ABB RobotStudio station: Laboratorio1Ruiz.rspag

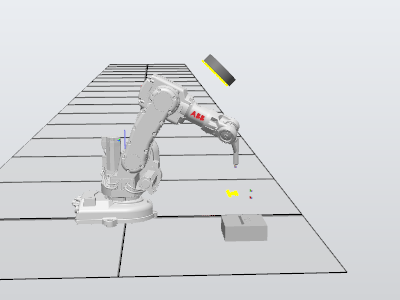
--- station ---
Station Laboratorio1 (saved by RobotStudio 25.5.11605.0)
Controller IRB140_6_81
  mechanical unit ROB_1: IRB140_6_81_C_03, 6 joints, base frame (0, 0, 0) mm
Layout (positions relative to the parent item):
  - IRB140_6_81_C_03 [mechanism, from %ABB.RobotStudio.Models.IRB140%\IRB140_6_81_C_G_03.rslib] at (0, 0, 0) mm; joint values [-0.1334, 0.4721, -0.017, 0.5827, 0.9537, -1.4192] (rad or m)
  - ToolLab1AlexaReyes [mechanism] at (588.01, -49.46, 449.3) mm, rotated rx 180 ry 30 rz -123.8 deg
      TCP ToolLab1AlexaReyes at (38.82, 1.24, 164.3) mm, rotated rx 0 ry 30 rz 0 deg
      links: Tool_3
  - Trayectorias2 [part] at (589.46, -613.7, 102.2) mm, rotated rx 0 ry 0 rz -90 deg, size 210 x 200 x 73 mm
  - Pieza_1 [part] at (-200, 0, 100) mm, rotated rx 0 ry 45 rz 0 deg, size 200 x 198.9 x 50 mm
  - SmartComponent_1 [smart component]
      signals: DI DI_04
      connections:
        LinearMover2.Executed -> LogicSRLatch.Reset
        LinearMover2.Executing -> LogicSRLatch.Set
        SmartComponent_1.DI_04 -> LinearMover2.Execute
    - LinearMover2 [smart component, from Components\LinearMover2.rslib]
        properties: Object=Trayectorias2; Direction=[0 0.001 0]; Distance=0.605; Duration=4.2; Reference=Global; ReferenceObject=(none)
  - SmartComponent_2 [smart component]
      signals: DI DI_05
      connections:
        SmartComponent_2.DI_05 -> LinearMover2_3.Execute
    - LinearMover2_3 [smart component, from Components\LinearMover2.rslib]
        properties: Object=Trayectorias2; Direction=[0 0.001 0]; Distance=0.605; Duration=4.2; Reference=Global; ReferenceObject=(none)
  - SmartComponent_3 [smart component]
      signals: DI DI_06
      connections:
        SmartComponent_3.DI_06 -> LinearMover2_5.Execute
    - LinearMover2_5 [smart component, from Components\LinearMover2.rslib]
        properties: Object=Trayectorias2; Direction=[0 -0.001 0]; Distance=1.21; Duration=8.4; Reference=Global; ReferenceObject=(none)
Attachment: ToolLab1AlexaReyes is attached to IRB140_6_81_C_03 / Link6
Station logic (signal -> signal, property => property):
  IRB140_6_81.DO_01 -> SmartComponent_1.DI_04
  IRB140_6_81.DO_02 -> SmartComponent_2.DI_05
  IRB140_6_81.DO_03 -> SmartComponent_3.DI_06

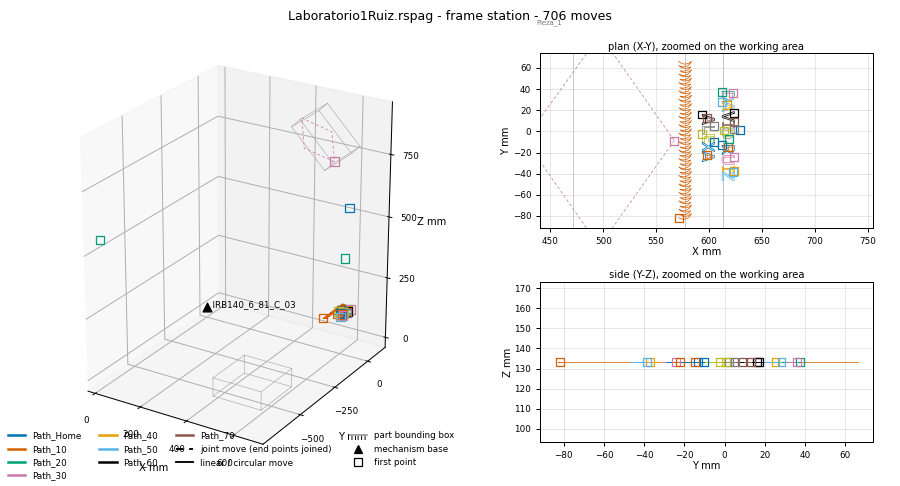
[picture p0: tool path of Laboratorio1Ruiz.rspag in frame station, 706 of 706 moves have a stored position in this frame; points joined in program order, loops and branches not executed]
--- Controller Data/IRB140_6_81/RAPID/TASK1/PROGMOD/Module1.mod ---
MODULE Module1
    PERS tooldata ToolLab1AlexaReyes:=[TRUE,[[38.819,1.24,164.297],[0.965925826,0,0.258819045,0]],[1,[0,0,1],[1,0,0,0],0,0,0]]; !CALIBRACIÓN VIRTUAL
    !PERS tooldata ToolLab1AlexaReyes:=[TRUE,[[37.2018,0.567088,156.366],[1,0,0,0]],[1,[0,0,0],[1,0,0,0],0,0,0]]; !CALIBRACIÓN FÍSICA
    CONST robtarget Target_Home:=[[629.167524851,1.24,563.73325724],[0.258819038,0,0.965925828,0],[0,-1,0,0],[9E+09,9E+09,9E+09,9E+09,9E+09,9E+09]];
    CONST robtarget Target_10:=[[118,32,0],[0.882142515,0,0,-0.470982573],[0,0,0,0],[9E+09,9E+09,9E+09,9E+09,9E+09,9E+09]];
    CONST robtarget Target_20:=[[115.336324555,30.849749419,0],[0.882142515,0,0,-0.470982573],[0,0,0,0],[9E+09,9E+09,9E+09,9E+09,9E+09,9E+09]];
    CONST robtarget Target_30:=[[112.437578714,30.725186884,0],[0.882142515,0,0,-0.470982573],[0,0,0,0],[9E+09,9E+09,9E+09,9E+09,9E+09,9E+09]];
    CONST robtarget Target_40:=[[109.685049159,31.642696736,0],[0.882142515,0,0,-0.470982573],[0,0,0,0],[9E+09,9E+09,9E+09,9E+09,9E+09,9E+09]];
    CONST robtarget Target_50:=[[107.440790007,33.481594268,0],[0.882142515,0,0,-0.470982573],[0,0,0,0],[9E+09,9E+09,9E+09,9E+09,9E+09,9E+09]];
    CONST robtarget Target_60:=[[106,36,0],[0.882142515,0,0,-0.470982573],[0,0,0,0],[9E+09,9E+09,9E+09,9E+09,9E+09,9E+09]];
    CONST robtarget Target_70:=[[108.368741055,34.163111606,0],[0.882142515,0,0,-0.470982573],[0,0,0,0],[9E+09,9E+09,9E+09,9E+09,9E+09,9E+09]];
    CONST robtarget Target_80:=[[111.247282109,33.326992858,0],[0.882142515,0,0,-0.470982573],[0,0,0,0],[9E+09,9E+09,9E+09,9E+09,9E+09,9E+09]];
    CONST robtarget Target_90:=[[114.231498793,33.609028207,0],[0.882142515,0,0,-0.470982573],[0,0,0,0],[9E+09,9E+09,9E+09,9E+09,9E+09,9E+09]];
    CONST robtarget Target_100:=[[116.902430719,34.969622123,0],[0.882142515,0,0,-0.470982573],[0,0,0,0],[9E+09,9E+09,9E+09,9E+09,9E+09,9E+09]];
    CONST robtarget Target_110:=[[113.892645843,34.654955892,0],[0.882142515,0,0,-0.470982573],[0,0,0,0],[9E+09,9E+09,9E+09,9E+09,9E+09,9E+09]];
    CONST robtarget Target_120:=[[111.01937121,35.058113631,0],[0.882142515,0,0,-0.470982573],[0,0,0,0],[9E+09,9E+09,9E+09,9E+09,9E+09,9E+09]];
    CONST robtarget Target_130:=[[108.478856861,36.459552219,0],[0.882142515,0,0,-0.470982573],[0,0,0,0],[9E+09,9E+09,9E+09,9E+09,9E+09,9E+09]];
    CONST robtarget Target_140:=[[106.60526948,38.674933361,0],[0.882142515,0,0,-0.470982573],[0,0,0,0],[9E+09,9E+09,9E+09,9E+09,9E+09,9E+09]];
    CONST robtarget Target_150:=[[109.768501207,37.609028207,0],[0.882142515,0,0,-0.470982573],[0,0,0,0],[9E+09,9E+09,9E+09,9E+09,9E+09,9E+09]];
    CONST robtarget Target_160:=[[112.752717891,37.326992858,0],[0.882142515,0,0,-0.470982573],[0,0,0,0],[9E+09,9E+09,9E+09,9E+09,9E+09,9E+09]];
    CONST robtarget Target_170:=[[115.631258945,38.163111606,0],[0.882142515,0,0,-0.470982573],[0,0,0,0],[9E+09,9E+09,9E+09,9E+09,9E+09,9E+09]];
    CONST robtarget Target_180:=[[118,40,0],[0.882142515,0,0,-0.470982573],[0,0,0,0],[9E+09,9E+09,9E+09,9E+09,9E+09,9E+09]];
    CONST robtarget Target_190:=[[115.336324555,38.849749419,0],[0.882142515,0,0,-0.470982573],[0,0,0,0],[9E+09,9E+09,9E+09,9E+09,9E+09,9E+09]];
    CONST robtarget Target_200:=[[112.437578714,38.725186884,0],[0.882142515,0,0,-0.470982573],[0,0,0,0],[9E+09,9E+09,9E+09,9E+09,9E+09,9E+09]];
    CONST robtarget Target_210:=[[109.685049159,39.642696736,0],[0.882142515,0,0,-0.470982573],[0,0,0,0],[9E+09,9E+09,9E+09,9E+09,9E+09,9E+09]];
    CONST robtarget Target_220:=[[107.440790007,41.481594268,0],[0.882142515,0,0,-0.470982573],[0,0,0,0],[9E+09,9E+09,9E+09,9E+09,9E+09,9E+09]];
    CONST robtarget Target_230:=[[106,44,0],[0.882142515,0,0,-0.470982573],[0,0,0,0],[9E+09,9E+09,9E+09,9E+09,9E+09,9E+09]];
    CONST robtarget Target_240:=[[108.368741055,42.163111606,0],[0.882142515,0,0,-0.470982573],[0,0,0,0],[9E+09,9E+09,9E+09,9E+09,9E+09,9E+09]];
    CONST robtarget Target_250:=[[111.247282109,41.326992858,0],[0.882142515,0,0,-0.470982573],[0,0,0,0],[9E+09,9E+09,9E+09,9E+09,9E+09,9E+09]];
    CONST robtarget Target_260:=[[114.231498793,41.609028207,0],[0.882142515,0,0,-0.470982573],[0,0,0,0],[9E+09,9E+09,9E+09,9E+09,9E+09,9E+09]];
    CONST robtarget Target_270:=[[116.902430719,42.969622123,0],[0.882142515,0,0,-0.470982573],[0,0,0,0],[9E+09,9E+09,9E+09,9E+09,9E+09,9E+09]];
    CONST robtarget Target_280:=[[113.892645843,42.654955892,0],[0.882142515,0,0,-0.470982573],[0,0,0,0],[9E+09,9E+09,9E+09,9E+09,9E+09,9E+09]];
    CONST robtarget Target_290:=[[111.01937121,43.058113631,0],[0.882142515,0,0,-0.470982573],[0,0,0,0],[9E+09,9E+09,9E+09,9E+09,9E+09,9E+09]];
    CONST robtarget Target_300:=[[108.478856861,44.459552219,0],[0.882142515,0,0,-0.470982573],[0,0,0,0],[9E+09,9E+09,9E+09,9E+09,9E+09,9E+09]];
    CONST robtarget Target_310:=[[106.60526948,46.674933361,0],[0.882142515,0,0,-0.470982573],[0,0,0,0],[9E+09,9E+09,9E+09,9E+09,9E+09,9E+09]];
    CONST robtarget Target_320:=[[109.768501207,45.609028207,0],[0.882142515,0,0,-0.470982573],[0,0,0,0],[9E+09,9E+09,9E+09,9E+09,9E+09,9E+09]];
    CONST robtarget Target_330:=[[112.752717891,45.326992858,0],[0.882142515,0,0,-0.470982573],[0,0,0,0],[9E+09,9E+09,9E+09,9E+09,9E+09,9E+09]];
    CONST robtarget Target_340:=[[115.631258945,46.163111606,0],[0.882142515,0,0,-0.470982573],[0,0,0,0],[9E+09,9E+09,9E+09,9E+09,9E+09,9E+09]];
    CONST robtarget Target_350:=[[118,48,0],[0.882142515,0,0,-0.470982573],[0,0,0,0],[9E+09,9E+09,9E+09,9E+09,9E+09,9E+09]];
    CONST robtarget Target_360:=[[115.336324555,46.849749419,0],[0.882142515,0,0,-0.470982573],[0,0,0,0],[9E+09,9E+09,9E+09,9E+09,9E+09,9E+09]];
    CONST robtarget Target_370:=[[112.437578714,46.725186884,0],[0.882142515,0,0,-0.470982573],[0,0,0,0],[9E+09,9E+09,9E+09,9E+09,9E+09,9E+09]];
    CONST robtarget Target_380:=[[109.685049159,47.642696736,0],[0.882142515,0,0,-0.470982573],[0,0,0,0],[9E+09,9E+09,9E+09,9E+09,9E+09,9E+09]];
    CONST robtarget Target_390:=[[107.440790007,49.481594268,0],[0.882142515,0,0,-0.470982573],[0,0,0,0],[9E+09,9E+09,9E+09,9E+09,9E+09,9E+09]];
    CONST robtarget Target_400:=[[106,52,0],[0.882142515,0,0,-0.470982573],[0,0,0,0],[9E+09,9E+09,9E+09,9E+09,9E+09,9E+09]];
    CONST robtarget Target_410:=[[108.368741055,50.163111606,0],[0.882142515,0,0,-0.470982573],[0,0,0,0],[9E+09,9E+09,9E+09,9E+09,9E+09,9E+09]];
    CONST robtarget Target_420:=[[111.247282109,49.326992858,0],[0.882142515,0,0,-0.470982573],[0,0,0,0],[9E+09,9E+09,9E+09,9E+09,9E+09,9E+09]];
    CONST robtarget Target_430:=[[114.231498793,49.609028207,0],[0.882142515,0,0,-0.470982573],[0,0,0,0],[9E+09,9E+09,9E+09,9E+09,9E+09,9E+09]];
    CONST robtarget Target_440:=[[116.902430719,50.969622123,0],[0.882142515,0,0,-0.470982573],[0,0,0,0],[9E+09,9E+09,9E+09,9E+09,9E+09,9E+09]];
    CONST robtarget Target_450:=[[113.892645843,50.654955892,0],[0.882142515,0,0,-0.470982573],[0,0,0,0],[9E+09,9E+09,9E+09,9E+09,9E+09,9E+09]];
    CONST robtarget Target_460:=[[111.01937121,51.058113631,0],[0.882142515,0,0,-0.470982573],[0,0,0,0],[9E+09,9E+09,9E+09,9E+09,9E+09,9E+09]];
    CONST robtarget Target_470:=[[108.478856861,52.459552219,0],[0.882142515,0,0,-0.470982573],[0,0,0,0],[9E+09,9E+09,9E+09,9E+09,9E+09,9E+09]];
    CONST robtarget Target_480:=[[106.60526948,54.674933361,0],[0.882142515,0,0,-0.470982573],[0,0,0,0],[9E+09,9E+09,9E+09,9E+09,9E+09,9E+09]];
    CONST robtarget Target_490:=[[109.768501207,53.609028207,0],[0.882142515,0,0,-0.470982573],[0,0,0,0],[9E+09,9E+09,9E+09,9E+09,9E+09,9E+09]];
    CONST robtarget Target_500:=[[112.752717891,53.326992858,0],[0.882142515,0,0,-0.470982573],[0,0,0,0],[9E+09,9E+09,9E+09,9E+09,9E+09,9E+09]];
    CONST robtarget Target_510:=[[115.631258945,54.163111606,0],[0.882142515,0,0,-0.470982573],[0,0,0,0],[9E+09,9E+09,9E+09,9E+09,9E+09,9E+09]];
    CONST robtarget Target_520:=[[118,56,0],[0.882142515,0,0,-0.470982573],[0,0,0,0],[9E+09,9E+09,9E+09,9E+09,9E+09,9E+09]];
    CONST robtarget Target_530:=[[115.336324555,54.849749419,0],[0.882142515,0,0,-0.470982573],[0,0,0,0],[9E+09,9E+09,9E+09,9E+09,9E+09,9E+09]];
    CONST robtarget Target_540:=[[112.437578714,54.725186884,0],[0.882142515,0,0,-0.470982573],[0,0,0,0],[9E+09,9E+09,9E+09,9E+09,9E+09,9E+09]];
    CONST robtarget Target_550:=[[109.685049159,55.642696736,0],[0.882142515,0,0,-0.470982573],[0,0,0,0],[9E+09,9E+09,9E+09,9E+09,9E+09,9E+09]];
    CONST robtarget Target_560:=[[107.440790007,57.481594268,0],[0.882142515,0,0,-0.470982573],[0,0,0,0],[9E+09,9E+09,9E+09,9E+09,9E+09,9E+09]];
    CONST robtarget Target_570:=[[106,60,0],[0.882142515,0,0,-0.470982573],[0,0,0,0],[9E+09,9E+09,9E+09,9E+09,9E+09,9E+09]];
    CONST robtarget Target_580:=[[108.368741055,58.163111606,0],[0.882142515,0,0,-0.470982573],[0,0,0,0],[9E+09,9E+09,9E+09,9E+09,9E+09,9E+09]];
    CONST robtarget Target_590:=[[111.247282109,57.326992858,0],[0.882142515,0,0,-0.470982573],[0,0,0,0],[9E+09,9E+09,9E+09,9E+09,9E+09,9E+09]];
    CONST robtarget Target_600:=[[114.231498793,57.609028207,0],[0.882142515,0,0,-0.470982573],[0,0,0,0],[9E+09,9E+09,9E+09,9E+09,9E+09,9E+09]];
    CONST robtarget Target_610:=[[116.902430719,58.969622123,0],[0.882142515,0,0,-0.470982573],[0,0,0,0],[9E+09,9E+09,9E+09,9E+09,9E+09,9E+09]];
    CONST robtarget Target_620:=[[113.892645843,58.654955892,0],[0.882142515,0,0,-0.470982573],[0,0,0,0],[9E+09,9E+09,9E+09,9E+09,9E+09,9E+09]];
    CONST robtarget Target_630:=[[111.01937121,59.058113631,0],[0.882142515,0,0,-0.470982573],[0,0,0,0],[9E+09,9E+09,9E+09,9E+09,9E+09,9E+09]];
    CONST robtarget Target_640:=[[108.478856861,60.459552219,0],[0.882142515,0,0,-0.470982573],[0,0,0,0],[9E+09,9E+09,9E+09,9E+09,9E+09,9E+09]];
    CONST robtarget Target_650:=[[106.60526948,62.674933361,0],[0.882142515,0,0,-0.470982573],[0,0,0,0],[9E+09,9E+09,9E+09,9E+09,9E+09,9E+09]];
    CONST robtarget Target_660:=[[109.768501207,61.609028207,0],[0.882142515,0,0,-0.470982573],[0,0,0,0],[9E+09,9E+09,9E+09,9E+09,9E+09,9E+09]];
    CONST robtarget Target_670:=[[112.752717891,61.326992858,0],[0.882142515,0,0,-0.470982573],[0,0,0,0],[9E+09,9E+09,9E+09,9E+09,9E+09,9E+09]];
    CONST robtarget Target_680:=[[115.631258945,62.163111606,0],[0.882142515,0,0,-0.470982573],[0,0,0,0],[9E+09,9E+09,9E+09,9E+09,9E+09,9E+09]];
    CONST robtarget Target_690:=[[118,64,0],[0.882142515,0,0,-0.470982573],[0,0,0,0],[9E+09,9E+09,9E+09,9E+09,9E+09,9E+09]];
    CONST robtarget Target_700:=[[115.336324555,62.849749419,0],[0.882142515,0,0,-0.470982573],[0,0,0,0],[9E+09,9E+09,9E+09,9E+09,9E+09,9E+09]];
    CONST robtarget Target_710:=[[112.437578714,62.725186884,0],[0.882142515,0,0,-0.470982573],[0,0,0,0],[9E+09,9E+09,9E+09,9E+09,9E+09,9E+09]];
    CONST robtarget Target_720:=[[109.685049159,63.642696736,0],[0.882142515,0,0,-0.470982573],[0,0,0,0],[9E+09,9E+09,9E+09,9E+09,9E+09,9E+09]];
    CONST robtarget Target_730:=[[107.440790007,65.481594268,0],[0.882142515,0,0,-0.470982573],[0,0,0,0],[9E+09,9E+09,9E+09,9E+09,9E+09,9E+09]];
    CONST robtarget Target_740:=[[106,68,0],[0.882142515,0,0,-0.470982573],[0,0,0,0],[9E+09,9E+09,9E+09,9E+09,9E+09,9E+09]];
    CONST robtarget Target_750:=[[108.368741055,66.163111606,0],[0.882142515,0,0,-0.470982573],[0,0,0,0],[9E+09,9E+09,9E+09,9E+09,9E+09,9E+09]];
    CONST robtarget Target_760:=[[111.247282109,65.326992858,0],[0.882142515,0,0,-0.470982573],[0,0,0,0],[9E+09,9E+09,9E+09,9E+09,9E+09,9E+09]];
    CONST robtarget Target_770:=[[114.231498793,65.609028207,0],[0.882142515,0,0,-0.470982573],[0,0,0,0],[9E+09,9E+09,9E+09,9E+09,9E+09,9E+09]];
    CONST robtarget Target_780:=[[116.902430719,66.969622123,0],[0.882142515,0,0,-0.470982573],[0,0,0,0],[9E+09,9E+09,9E+09,9E+09,9E+09,9E+09]];
    CONST robtarget Target_790:=[[113.892645843,66.654955892,0],[0.882142515,0,0,-0.470982573],[0,0,0,0],[9E+09,9E+09,9E+09,9E+09,9E+09,9E+09]];
    CONST robtarget Target_800:=[[111.01937121,67.058113631,0],[0.882142515,0,0,-0.470982573],[0,0,0,0],[9E+09,9E+09,9E+09,9E+09,9E+09,9E+09]];
    CONST robtarget Target_810:=[[108.478856861,68.459552219,0],[0.882142515,0,0,-0.470982573],[0,0,0,0],[9E+09,9E+09,9E+09,9E+09,9E+09,9E+09]];
    CONST robtarget Target_820:=[[106.60526948,70.674933361,0],[0.882142515,0,0,-0.470982573],[0,0,0,0],[9E+09,9E+09,9E+09,9E+09,9E+09,9E+09]];
    CONST robtarget Target_830:=[[109.768501207,69.609028207,0],[0.882142515,0,0,-0.470982573],[0,0,0,0],[9E+09,9E+09,9E+09,9E+09,9E+09,9E+09]];
    CONST robtarget Target_840:=[[112.752717891,69.326992858,0],[0.882142515,0,0,-0.470982573],[0,0,0,0],[9E+09,9E+09,9E+09,9E+09,9E+09,9E+09]];
    CONST robtarget Target_850:=[[115.631258945,70.163111606,0],[0.882142515,0,0,-0.470982573],[0,0,0,0],[9E+09,9E+09,9E+09,9E+09,9E+09,9E+09]];
    CONST robtarget Target_860:=[[118,72,0],[0.882142515,0,0,-0.470982573],[0,0,0,0],[9E+09,9E+09,9E+09,9E+09,9E+09,9E+09]];
    CONST robtarget Target_870:=[[115.336324555,70.849749419,0],[0.882142515,0,0,-0.470982573],[0,0,0,0],[9E+09,9E+09,9E+09,9E+09,9E+09,9E+09]];
    CONST robtarget Target_880:=[[112.437578714,70.725186884,0],[0.882142515,0,0,-0.470982573],[0,0,0,0],[9E+09,9E+09,9E+09,9E+09,9E+09,9E+09]];
    CONST robtarget Target_890:=[[109.685049159,71.642696736,0],[0.882142515,0,0,-0.470982573],[0,0,0,0],[9E+09,9E+09,9E+09,9E+09,9E+09,9E+09]];
    CONST robtarget Target_900:=[[107.440790007,73.481594268,0],[0.882142515,0,0,-0.470982573],[0,0,0,0],[9E+09,9E+09,9E+09,9E+09,9E+09,9E+09]];
    CONST robtarget Target_910:=[[106,76,0],[0.882142515,0,0,-0.470982573],[0,0,0,0],[9E+09,9E+09,9E+09,9E+09,9E+09,9E+09]];
    CONST robtarget Target_920:=[[108.368741055,74.163111606,0],[0.882142515,0,0,-0.470982573],[0,0,0,0],[9E+09,9E+09,9E+09,9E+09,9E+09,9E+09]];
    CONST robtarget Target_930:=[[111.247282109,73.326992858,0],[0.882142515,0,0,-0.470982573],[0,0,0,0],[9E+09,9E+09,9E+09,9E+09,9E+09,9E+09]];
    CONST robtarget Target_940:=[[114.231498793,73.609028207,0],[0.882142515,0,0,-0.470982573],[0,0,0,0],[9E+09,9E+09,9E+09,9E+09,9E+09,9E+09]];
    CONST robtarget Target_950:=[[116.902430719,74.969622123,0],[0.882142515,0,0,-0.470982573],[0,0,0,0],[9E+09,9E+09,9E+09,9E+09,9E+09,9E+09]];
    CONST robtarget Target_960:=[[113.892645843,74.654955892,0],[0.882142515,0,0,-0.470982573],[0,0,0,0],[9E+09,9E+09,9E+09,9E+09,9E+09,9E+09]];
    CONST robtarget Target_970:=[[111.01937121,75.058113631,0],[0.882142515,0,0,-0.470982573],[0,0,0,0],[9E+09,9E+09,9E+09,9E+09,9E+09,9E+09]];
    CONST robtarget Target_980:=[[108.478856861,76.459552219,0],[0.882142515,0,0,-0.470982573],[0,0,0,0],[9E+09,9E+09,9E+09,9E+09,9E+09,9E+09]];
    CONST robtarget Target_990:=[[106.60526948,78.674933361,0],[0.882142515,0,0,-0.470982573],[0,0,0,0],[9E+09,9E+09,9E+09,9E+09,9E+09,9E+09]];
    CONST robtarget Target_1000:=[[109.768501207,77.609028207,0],[0.882142515,0,0,-0.470982573],[0,0,0,0],[9E+09,9E+09,9E+09,9E+09,9E+09,9E+09]];
    CONST robtarget Target_1010:=[[112.752717891,77.326992858,0],[0.882142515,0,0,-0.470982573],[0,0,0,0],[9E+09,9E+09,9E+09,9E+09,9E+09,9E+09]];
    CONST robtarget Target_1020:=[[115.631258945,78.163111606,0],[0.882142515,0,0,-0.470982573],[0,0,0,0],[9E+09,9E+09,9E+09,9E+09,9E+09,9E+09]];
    CONST robtarget Target_1030:=[[118,80,0],[0.882142515,0,0,-0.470982573],[0,0,0,0],[9E+09,9E+09,9E+09,9E+09,9E+09,9E+09]];
    CONST robtarget Target_1040:=[[115.336324555,78.849749419,0],[0.882142515,0,0,-0.470982573],[0,0,0,0],[9E+09,9E+09,9E+09,9E+09,9E+09,9E+09]];
    CONST robtarget Target_1050:=[[112.437578714,78.725186884,0],[0.882142515,0,0,-0.470982573],[0,0,0,0],[9E+09,9E+09,9E+09,9E+09,9E+09,9E+09]];
    CONST robtarget Target_1060:=[[109.685049159,79.642696736,0],[0.882142515,0,0,-0.470982573],[0,0,0,0],[9E+09,9E+09,9E+09,9E+09,9E+09,9E+09]];
    CONST robtarget Target_1070:=[[107.440790007,81.481594268,0],[0.882142515,0,0,-0.470982573],[0,0,0,0],[9E+09,9E+09,9E+09,9E+09,9E+09,9E+09]];
    CONST robtarget Target_1080:=[[106,84,0],[0.882142515,0,0,-0.470982573],[0,0,0,0],[9E+09,9E+09,9E+09,9E+09,9E+09,9E+09]];
    CONST robtarget Target_1090:=[[108.368741055,82.163111606,0],[0.882142515,0,0,-0.470982573],[0,0,0,0],[9E+09,9E+09,9E+09,9E+09,9E+09,9E+09]];
    CONST robtarget Target_1100:=[[111.247282109,81.326992858,0],[0.882142515,0,0,-0.470982573],[0,0,0,0],[9E+09,9E+09,9E+09,9E+09,9E+09,9E+09]];
    CONST robtarget Target_1110:=[[114.231498793,81.609028207,0],[0.882142515,0,0,-0.470982573],[0,0,0,0],[9E+09,9E+09,9E+09,9E+09,9E+09,9E+09]];
    CONST robtarget Target_1120:=[[116.902430719,82.969622123,0],[0.882142515,0,0,-0.470982573],[0,0,0,0],[9E+09,9E+09,9E+09,9E+09,9E+09,9E+09]];
    CONST robtarget Target_1130:=[[113.892645843,82.654955892,0],[0.882142515,0,0,-0.470982573],[0,0,0,0],[9E+09,9E+09,9E+09,9E+09,9E+09,9E+09]];
    CONST robtarget Target_1140:=[[111.01937121,83.058113631,0],[0.882142515,0,0,-0.470982573],[0,0,0,0],[9E+09,9E+09,9E+09,9E+09,9E+09,9E+09]];
    CONST robtarget Target_1150:=[[108.478856861,84.459552219,0],[0.882142515,0,0,-0.470982573],[0,0,0,0],[9E+09,9E+09,9E+09,9E+09,9E+09,9E+09]];
    CONST robtarget Target_1160:=[[106.60526948,86.674933361,0],[0.882142515,0,0,-0.470982573],[0,0,0,0],[9E+09,9E+09,9E+09,9E+09,9E+09,9E+09]];
    CONST robtarget Target_1170:=[[109.768501207,85.609028207,0],[0.882142515,0,0,-0.470982573],[0,0,0,0],[9E+09,9E+09,9E+09,9E+09,9E+09,9E+09]];
    CONST robtarget Target_1180:=[[112.752717891,85.326992858,0],[0.882142515,0,0,-0.470982573],[0,0,0,0],[9E+09,9E+09,9E+09,9E+09,9E+09,9E+09]];
    CONST robtarget Target_1190:=[[115.631258945,86.163111606,0],[0.882142515,0,0,-0.470982573],[0,0,0,0],[9E+09,9E+09,9E+09,9E+09,9E+09,9E+09]];
    CONST robtarget Target_1200:=[[118,88,0],[0.882142515,0,0,-0.470982573],[0,0,0,0],[9E+09,9E+09,9E+09,9E+09,9E+09,9E+09]];
    CONST robtarget Target_1210:=[[115.336324555,86.849749419,0],[0.882142515,0,0,-0.470982573],[0,0,0,0],[9E+09,9E+09,9E+09,9E+09,9E+09,9E+09]];
    CONST robtarget Target_1220:=[[112.437578714,86.725186884,0],[0.882142515,0,0,-0.470982573],[0,0,0,0],[9E+09,9E+09,9E+09,9E+09,9E+09,9E+09]];
    CONST robtarget Target_1230:=[[109.685049159,87.642696736,0],[0.882142515,0,0,-0.470982573],[0,0,0,0],[9E+09,9E+09,9E+09,9E+09,9E+09,9E+09]];
    CONST robtarget Target_1240:=[[107.440790007,89.481594268,0],[0.882142515,0,0,-0.470982573],[0,0,0,0],[9E+09,9E+09,9E+09,9E+09,9E+09,9E+09]];
    CONST robtarget Target_1250:=[[106,92,0],[0.882142515,0,0,-0.470982573],[0,0,0,0],[9E+09,9E+09,9E+09,9E+09,9E+09,9E+09]];
    CONST robtarget Target_1260:=[[108.368741055,90.163111606,0],[0.882142515,0,0,-0.470982573],[0,0,0,0],[9E+09,9E+09,9E+09,9E+09,9E+09,9E+09]];
    CONST robtarget Target_1270:=[[111.247282109,89.326992858,0],[0.882142515,0,0,-0.470982573],[0,0,0,0],[9E+09,9E+09,9E+09,9E+09,9E+09,9E+09]];
    CONST robtarget Target_1280:=[[114.231498793,89.609028207,0],[0.882142515,0,0,-0.470982573],[0,0,0,0],[9E+09,9E+09,9E+09,9E+09,9E+09,9E+09]];
    CONST robtarget Target_1290:=[[116.902430719,90.969622123,0],[0.882142515,0,0,-0.470982573],[0,0,0,0],[9E+09,9E+09,9E+09,9E+09,9E+09,9E+09]];
    CONST robtarget Target_1300:=[[113.892645843,90.654955892,0],[0.882142515,0,0,-0.470982573],[0,0,0,0],[9E+09,9E+09,9E+09,9E+09,9E+09,9E+09]];
    CONST robtarget Target_1310:=[[111.01937121,91.058113631,0],[0.882142515,0,0,-0.470982573],[0,0,0,0],[9E+09,9E+09,9E+09,9E+09,9E+09,9E+09]];
    CONST robtarget Target_1320:=[[108.478856861,92.459552219,0],[0.882142515,0,0,-0.470982573],[0,0,0,0],[9E+09,9E+09,9E+09,9E+09,9E+09,9E+09]];
    CONST robtarget Target_1330:=[[106.60526948,94.674933361,0],[0.882142515,0,0,-0.470982573],[0,0,0,0],[9E+09,9E+09,9E+09,9E+09,9E+09,9E+09]];
    CONST robtarget Target_1340:=[[109.768501207,93.609028207,0],[0.882142515,0,0,-0.470982573],[0,0,0,0],[9E+09,9E+09,9E+09,9E+09,9E+09,9E+09]];
    CONST robtarget Target_1350:=[[112.752717891,93.326992858,0],[0.882142515,0,0,-0.470982573],[0,0,0,0],[9E+09,9E+09,9E+09,9E+09,9E+09,9E+09]];
    CONST robtarget Target_1360:=[[115.631258945,94.163111606,0],[0.882142515,0,0,-0.470982573],[0,0,0,0],[9E+09,9E+09,9E+09,9E+09,9E+09,9E+09]];
    CONST robtarget Target_1370:=[[118,96,0],[0.882142515,0,0,-0.470982573],[0,0,0,0],[9E+09,9E+09,9E+09,9E+09,9E+09,9E+09]];
    CONST robtarget Target_1380:=[[115.336324555,94.849749419,0],[0.882142515,0,0,-0.470982573],[0,0,0,0],[9E+09,9E+09,9E+09,9E+09,9E+09,9E+09]];
    CONST robtarget Target_1390:=[[112.437578714,94.725186884,0],[0.882142515,0,0,-0.470982573],[0,0,0,0],[9E+09,9E+09,9E+09,9E+09,9E+09,9E+09]];
    CONST robtarget Target_1400:=[[109.685049159,95.642696736,0],[0.882142515,0,0,-0.470982573],[0,0,0,0],[9E+09,9E+09,9E+09,9E+09,9E+09,9E+09]];
    CONST robtarget Target_1410:=[[107.440790007,97.481594268,0],[0.882142515,0,0,-0.470982573],[0,0,0,0],[9E+09,9E+09,9E+09,9E+09,9E+09,9E+09]];
    CONST robtarget Target_1420:=[[106,100,0],[0.882142515,0,0,-0.470982573],[0,0,0,0],[9E+09,9E+09,9E+09,9E+09,9E+09,9E+09]];
    CONST robtarget Target_1430:=[[108.368741055,98.163111606,0],[0.882142515,0,0,-0.470982573],[0,0,0,0],[9E+09,9E+09,9E+09,9E+09,9E+09,9E+09]];
    CONST robtarget Target_1440:=[[111.247282109,97.326992858,0],[0.882142515,0,0,-0.470982573],[0,0,0,0],[9E+09,9E+09,9E+09,9E+09,9E+09,9E+09]];
    CONST robtarget Target_1450:=[[114.231498793,97.609028207,0],[0.882142515,0,0,-0.470982573],[0,0,0,0],[9E+09,9E+09,9E+09,9E+09,9E+09,9E+09]];
    CONST robtarget Target_1460:=[[116.902430719,98.969622123,0],[0.882142515,0,0,-0.470982573],[0,0,0,0],[9E+09,9E+09,9E+09,9E+09,9E+09,9E+09]];
    CONST robtarget Target_1470:=[[113.892645843,98.654955892,0],[0.882142515,0,0,-0.470982573],[0,0,0,0],[9E+09,9E+09,9E+09,9E+09,9E+09,9E+09]];
    CONST robtarget Target_1480:=[[111.01937121,99.058113631,0],[0.882142515,0,0,-0.470982573],[0,0,0,0],[9E+09,9E+09,9E+09,9E+09,9E+09,9E+09]];
    CONST robtarget Target_1490:=[[108.478856861,100.459552219,0],[0.882142515,0,0,-0.470982573],[0,0,0,0],[9E+09,9E+09,9E+09,9E+09,9E+09,9E+09]];
    CONST robtarget Target_1500:=[[106.60526948,102.674933361,0],[0.882142515,0,0,-0.470982573],[0,0,0,0],[9E+09,9E+09,9E+09,9E+09,9E+09,9E+09]];
    CONST robtarget Target_1510:=[[109.768501207,101.609028207,0],[0.882142515,0,0,-0.470982573],[0,0,0,0],[9E+09,9E+09,9E+09,9E+09,9E+09,9E+09]];
    CONST robtarget Target_1520:=[[112.752717891,101.326992858,0],[0.882142515,0,0,-0.470982573],[0,0,0,0],[9E+09,9E+09,9E+09,9E+09,9E+09,9E+09]];
    TASK PERS wobjdata Workobject_1:=[FALSE,TRUE,"",[[689.46,-113.7,173.2],[0,-0.707106781,0.707106781,0]],[[0,0,40],[0.707106781,0,0,0.707106781]]];
    CONST robtarget Target_1530:=[[115.631258945,102.163111606,0],[0.882142515,0,0,-0.470982573],[0,0,0,0],[9E+09,9E+09,9E+09,9E+09,9E+09,9E+09]];
    CONST robtarget Target_1540:=[[118,104,0],[0.882142515,0,0,-0.470982573],[0,0,0,0],[9E+09,9E+09,9E+09,9E+09,9E+09,9E+09]];
    CONST robtarget Target_1550:=[[115.336324555,102.849749419,0],[0.882142515,0,0,-0.470982573],[0,0,0,0],[9E+09,9E+09,9E+09,9E+09,9E+09,9E+09]];
    CONST robtarget Target_1560:=[[112.437578714,102.725186884,0],[0.882142515,0,0,-0.470982573],[0,0,0,0],[9E+09,9E+09,9E+09,9E+09,9E+09,9E+09]];
    CONST robtarget Target_1570:=[[109.685049159,103.642696736,0],[0.882142515,0,0,-0.470982573],[0,0,0,0],[9E+09,9E+09,9E+09,9E+09,9E+09,9E+09]];
    CONST robtarget Target_1580:=[[107.440790007,105.481594268,0],[0.882142515,0,0,-0.470982573],[0,0,0,0],[9E+09,9E+09,9E+09,9E+09,9E+09,9E+09]];
    CONST robtarget Target_1590:=[[106,108,0],[0.882142515,0,0,-0.470982573],[0,0,0,0],[9E+09,9E+09,9E+09,9E+09,9E+09,9E+09]];
    CONST robtarget Target_1600:=[[108.368741055,106.163111606,0],[0.882142515,0,0,-0.470982573],[0,0,0,0],[9E+09,9E+09,9E+09,9E+09,9E+09,9E+09]];
    CONST robtarget Target_1610:=[[111.247282109,105.326992858,0],[0.882142515,0,0,-0.470982573],[0,0,0,0],[9E+09,9E+09,9E+09,9E+09,9E+09,9E+09]];
    CONST robtarget Target_1620:=[[114.231498793,105.609028207,0],[0.882142515,0,0,-0.470982573],[0,0,0,0],[9E+09,9E+09,9E+09,9E+09,9E+09,9E+09]];
    CONST robtarget Target_1630:=[[116.902430719,106.969622123,0],[0.882142515,0,0,-0.470982573],[0,0,0,0],[9E+09,9E+09,9E+09,9E+09,9E+09,9E+09]];
    CONST robtarget Target_1640:=[[113.892645843,106.654955892,0],[0.882142515,0,0,-0.470982573],[0,0,0,0],[9E+09,9E+09,9E+09,9E+09,9E+09,9E+09]];
    CONST robtarget Target_1650:=[[111.01937121,107.058113631,0],[0.882142515,0,0,-0.470982573],[0,0,0,0],[9E+09,9E+09,9E+09,9E+09,9E+09,9E+09]];
    CONST robtarget Target_1660:=[[108.478856861,108.459552219,0],[0.882142515,0,0,-0.470982573],[0,0,0,0],[9E+09,9E+09,9E+09,9E+09,9E+09,9E+09]];
    CONST robtarget Target_1670:=[[106.60526948,110.674933361,0],[0.882142515,0,0,-0.470982573],[0,0,0,0],[9E+09,9E+09,9E+09,9E+09,9E+09,9E+09]];
    CONST robtarget Target_1680:=[[109.768501207,109.609028207,0],[0.882142515,0,0,-0.470982573],[0,0,0,0],[9E+09,9E+09,9E+09,9E+09,9E+09,9E+09]];
    CONST robtarget Target_1690:=[[112.752717891,109.326992858,0],[0.882142515,0,0,-0.470982573],[0,0,0,0],[9E+09,9E+09,9E+09,9E+09,9E+09,9E+09]];
    CONST robtarget Target_1700:=[[115.631258945,110.163111606,0],[0.882142515,0,0,-0.470982573],[0,0,0,0],[9E+09,9E+09,9E+09,9E+09,9E+09,9E+09]];
    CONST robtarget Target_1710:=[[118,112,0],[0.882142515,0,0,-0.470982573],[0,0,0,0],[9E+09,9E+09,9E+09,9E+09,9E+09,9E+09]];
    CONST robtarget Target_1720:=[[115.336324555,110.849749419,0],[0.882142515,0,0,-0.470982573],[0,0,0,0],[9E+09,9E+09,9E+09,9E+09,9E+09,9E+09]];
    CONST robtarget Target_1730:=[[112.437578714,110.725186884,0],[0.882142515,0,0,-0.470982573],[0,0,0,0],[9E+09,9E+09,9E+09,9E+09,9E+09,9E+09]];
    CONST robtarget Target_1740:=[[109.685049159,111.642696736,0],[0.882142515,0,0,-0.470982573],[0,0,0,0],[9E+09,9E+09,9E+09,9E+09,9E+09,9E+09]];
    CONST robtarget Target_1750:=[[107.440790007,113.481594268,0],[0.882142515,0,0,-0.470982573],[0,0,0,0],[9E+09,9E+09,9E+09,9E+09,9E+09,9E+09]];
    CONST robtarget Target_1760:=[[106,116,0],[0.882142515,0,0,-0.470982573],[0,0,0,0],[9E+09,9E+09,9E+09,9E+09,9E+09,9E+09]];
    CONST robtarget Target_1770:=[[108.368741055,114.163111606,0],[0.882142515,0,0,-0.470982573],[0,0,0,0],[9E+09,9E+09,9E+09,9E+09,9E+09,9E+09]];
    CONST robtarget Target_1780:=[[111.247282109,113.326992858,0],[0.882142515,0,0,-0.470982573],[0,0,0,0],[9E+09,9E+09,9E+09,9E+09,9E+09,9E+09]];
    CONST robtarget Target_1790:=[[114.231498793,113.609028207,0],[0.882142515,0,0,-0.470982573],[0,0,0,0],[9E+09,9E+09,9E+09,9E+09,9E+09,9E+09]];
    CONST robtarget Target_1800:=[[116.902430719,114.969622123,0],[0.882142515,0,0,-0.470982573],[0,0,0,0],[9E+09,9E+09,9E+09,9E+09,9E+09,9E+09]];
    CONST robtarget Target_1810:=[[113.892645843,114.654955892,0],[0.882142515,0,0,-0.470982573],[0,0,0,0],[9E+09,9E+09,9E+09,9E+09,9E+09,9E+09]];
    CONST robtarget Target_1820:=[[111.01937121,115.058113631,0],[0.882142515,0,0,-0.470982573],[0,0,0,0],[9E+09,9E+09,9E+09,9E+09,9E+09,9E+09]];
    CONST robtarget Target_1830:=[[108.478856861,116.459552219,0],[0.882142515,0,0,-0.470982573],[0,0,0,0],[9E+09,9E+09,9E+09,9E+09,9E+09,9E+09]];
    CONST robtarget Target_1840:=[[106.60526948,118.674933361,0],[0.882142515,0,0,-0.470982573],[0,0,0,0],[9E+09,9E+09,9E+09,9E+09,9E+09,9E+09]];
    CONST robtarget Target_1850:=[[109.768501207,117.609028207,0],[0.882142515,0,0,-0.470982573],[0,0,0,0],[9E+09,9E+09,9E+09,9E+09,9E+09,9E+09]];
    CONST robtarget Target_1860:=[[112.752717891,117.326992858,0],[0.882142515,0,0,-0.470982573],[0,0,0,0],[9E+09,9E+09,9E+09,9E+09,9E+09,9E+09]];
    CONST robtarget Target_1870:=[[115.631258945,118.163111606,0],[0.882142515,0,0,-0.470982573],[0,0,0,0],[9E+09,9E+09,9E+09,9E+09,9E+09,9E+09]];
    CONST robtarget Target_1880:=[[118,120,0],[0.882142515,0,0,-0.470982573],[0,0,0,0],[9E+09,9E+09,9E+09,9E+09,9E+09,9E+09]];
    CONST robtarget Target_1890:=[[115.336324555,118.849749419,0],[0.882142515,0,0,-0.470982573],[0,0,0,0],[9E+09,9E+09,9E+09,9E+09,9E+09,9E+09]];
    CONST robtarget Target_1900:=[[112.437578714,118.725186884,0],[0.882142515,0,0,-0.470982573],[0,0,0,0],[9E+09,9E+09,9E+09,9E+09,9E+09,9E+09]];
    CONST robtarget Target_1910:=[[109.685049159,119.642696736,0],[0.882142515,0,0,-0.470982573],[0,0,0,0],[9E+09,9E+09,9E+09,9E+09,9E+09,9E+09]];
    CONST robtarget Target_1920:=[[107.440790007,121.481594268,0],[0.882142515,0,0,-0.470982573],[0,0,0,0],[9E+09,9E+09,9E+09,9E+09,9E+09,9E+09]];
    CONST robtarget Target_1930:=[[106,124,0],[0.882142515,0,0,-0.470982573],[0,0,0,0],[9E+09,9E+09,9E+09,9E+09,9E+09,9E+09]];
    CONST robtarget Target_1940:=[[108.368741055,122.163111606,0],[0.882142515,0,0,-0.470982573],[0,0,0,0],[9E+09,9E+09,9E+09,9E+09,9E+09,9E+09]];
    CONST robtarget Target_1950:=[[111.247282109,121.326992858,0],[0.882142515,0,0,-0.470982573],[0,0,0,0],[9E+09,9E+09,9E+09,9E+09,9E+09,9E+09]];
    CONST robtarget Target_1960:=[[114.231498793,121.609028207,0],[0.882142515,0,0,-0.470982573],[0,0,0,0],[9E+09,9E+09,9E+09,9E+09,9E+09,9E+09]];
    CONST robtarget Target_1970:=[[116.902430719,122.969622123,0],[0.882142515,0,0,-0.470982573],[0,0,0,0],[9E+09,9E+09,9E+09,9E+09,9E+09,9E+09]];
    CONST robtarget Target_1980:=[[113.892645843,122.654955892,0],[0.882142515,0,0,-0.470982573],[0,0,0,0],[9E+09,9E+09,9E+09,9E+09,9E+09,9E+09]];
    CONST robtarget Target_1990:=[[111.01937121,123.058113631,0],[0.882142515,0,0,-0.470982573],[0,0,0,0],[9E+09,9E+09,9E+09,9E+09,9E+09,9E+09]];
    CONST robtarget Target_2000:=[[108.478856861,124.459552219,0],[0.882142515,0,0,-0.470982573],[0,0,0,0],[9E+09,9E+09,9E+09,9E+09,9E+09,9E+09]];
    CONST robtarget Target_2010:=[[106.60526948,126.674933361,0],[0.882142515,0,0,-0.470982573],[0,0,0,0],[9E+09,9E+09,9E+09,9E+09,9E+09,9E+09]];
    CONST robtarget Target_2020:=[[109.768501207,125.609028207,0],[0.882142515,0,0,-0.470982573],[0,0,0,0],[9E+09,9E+09,9E+09,9E+09,9E+09,9E+09]];
    CONST robtarget Target_2030:=[[112.752717891,125.326992858,0],[0.882142515,0,0,-0.470982573],[0,0,0,0],[9E+09,9E+09,9E+09,9E+09,9E+09,9E+09]];
    CONST robtarget Target_2040:=[[115.631258945,126.163111606,0],[0.882142515,0,0,-0.470982573],[0,0,0,0],[9E+09,9E+09,9E+09,9E+09,9E+09,9E+09]];
    CONST robtarget Target_2050:=[[118,128,0],[0.882142515,0,0,-0.470982573],[0,0,0,0],[9E+09,9E+09,9E+09,9E+09,9E+09,9E+09]];
    CONST robtarget Target_2060:=[[115.336324555,126.849749419,0],[0.882142515,0,0,-0.470982573],[0,0,0,0],[9E+09,9E+09,9E+09,9E+09,9E+09,9E+09]];
    CONST robtarget Target_2070:=[[112.437578714,126.725186884,0],[0.882142515,0,0,-0.470982573],[0,0,0,0],[9E+09,9E+09,9E+09,9E+09,9E+09,9E+09]];
    CONST robtarget Target_2080:=[[109.685049159,127.642696736,0],[0.882142515,0,0,-0.470982573],[0,0,0,0],[9E+09,9E+09,9E+09,9E+09,9E+09,9E+09]];
    CONST robtarget Target_2090:=[[107.440790007,129.481594268,0],[0.882142515,0,0,-0.470982573],[0,0,0,0],[9E+09,9E+09,9E+09,9E+09,9E+09,9E+09]];
    CONST robtarget Target_2100:=[[106,132,0],[0.882142515,0,0,-0.470982573],[0,0,0,0],[9E+09,9E+09,9E+09,9E+09,9E+09,9E+09]];
    CONST robtarget Target_2110:=[[108.368741055,130.163111606,0],[0.882142515,0,0,-0.470982573],[0,0,0,0],[9E+09,9E+09,9E+09,9E+09,9E+09,9E+09]];
    CONST robtarget Target_2120:=[[111.247282109,129.326992858,0],[0.882142515,0,0,-0.470982573],[0,0,0,0],[9E+09,9E+09,9E+09,9E+09,9E+09,9E+09]];
    CONST robtarget Target_2130:=[[114.231498793,129.609028207,0],[0.882142515,0,0,-0.470982573],[0,0,0,0],[9E+09,9E+09,9E+09,9E+09,9E+09,9E+09]];
    CONST robtarget Target_2140:=[[116.902430719,130.969622123,0],[0.882142515,0,0,-0.470982573],[0,0,0,0],[9E+09,9E+09,9E+09,9E+09,9E+09,9E+09]];
    CONST robtarget Target_2150:=[[113.892645843,130.654955892,0],[0.882142515,0,0,-0.470982573],[0,0,0,0],[9E+09,9E+09,9E+09,9E+09,9E+09,9E+09]];
    CONST robtarget Target_2160:=[[111.01937121,131.058113631,0],[0.882142515,0,0,-0.470982573],[0,0,0,0],[9E+09,9E+09,9E+09,9E+09,9E+09,9E+09]];
    CONST robtarget Target_2170:=[[108.478856861,132.459552219,0],[0.882142515,0,0,-0.470982573],[0,0,0,0],[9E+09,9E+09,9E+09,9E+09,9E+09,9E+09]];
    CONST robtarget Target_2180:=[[106.60526948,134.674933361,0],[0.882142515,0,0,-0.470982573],[0,0,0,0],[9E+09,9E+09,9E+09,9E+09,9E+09,9E+09]];
    CONST robtarget Target_2190:=[[109.768501207,133.609028207,0],[0.882142515,0,0,-0.470982573],[0,0,0,0],[9E+09,9E+09,9E+09,9E+09,9E+09,9E+09]];
    CONST robtarget Target_2200:=[[112.752717891,133.326992858,0],[0.882142515,0,0,-0.470982573],[0,0,0,0],[9E+09,9E+09,9E+09,9E+09,9E+09,9E+09]];
    CONST robtarget Target_2210:=[[115.631258945,134.163111606,0],[0.882142515,0,0,-0.470982573],[0,0,0,0],[9E+09,9E+09,9E+09,9E+09,9E+09,9E+09]];
    CONST robtarget Target_2220:=[[118,136,0],[0.882142515,0,0,-0.470982573],[0,0,0,0],[9E+09,9E+09,9E+09,9E+09,9E+09,9E+09]];
    CONST robtarget Target_2230:=[[115.336324555,134.849749419,0],[0.882142515,0,0,-0.470982573],[0,0,0,0],[9E+09,9E+09,9E+09,9E+09,9E+09,9E+09]];
    CONST robtarget Target_2240:=[[112.437578714,134.725186884,0],[0.882142515,0,0,-0.470982573],[0,0,0,0],[9E+09,9E+09,9E+09,9E+09,9E+09,9E+09]];
    CONST robtarget Target_2250:=[[109.685049159,135.642696736,0],[0.882142515,0,0,-0.470982573],[0,0,0,0],[9E+09,9E+09,9E+09,9E+09,9E+09,9E+09]];
    CONST robtarget Target_2260:=[[107.440790007,137.481594268,0],[0.882142515,0,0,-0.470982573],[0,0,0,0],[9E+09,9E+09,9E+09,9E+09,9E+09,9E+09]];
    CONST robtarget Target_2270:=[[106,140,0],[0.882142515,0,0,-0.470982573],[0,0,0,0],[9E+09,9E+09,9E+09,9E+09,9E+09,9E+09]];
    CONST robtarget Target_2280:=[[108.368741055,138.163111606,0],[0.882142515,0,0,-0.470982573],[0,0,0,0],[9E+09,9E+09,9E+09,9E+09,9E+09,9E+09]];
    CONST robtarget Target_2290:=[[111.247282109,137.326992858,0],[0.882142515,0,0,-0.470982573],[0,0,0,0],[9E+09,9E+09,9E+09,9E+09,9E+09,9E+09]];
    CONST robtarget Target_2300:=[[114.231498793,137.609028207,0],[0.882142515,0,0,-0.470982573],[0,0,0,0],[9E+09,9E+09,9E+09,9E+09,9E+09,9E+09]];
    CONST robtarget Target_2310:=[[116.902430719,138.969622123,0],[0.882142515,0,0,-0.470982573],[0,0,0,0],[9E+09,9E+09,9E+09,9E+09,9E+09,9E+09]];
    CONST robtarget Target_2320:=[[113.892645843,138.654955892,0],[0.882142515,0,0,-0.470982573],[0,0,0,0],[9E+09,9E+09,9E+09,9E+09,9E+09,9E+09]];
    CONST robtarget Target_2330:=[[111.01937121,139.058113631,0],[0.882142515,0,0,-0.470982573],[0,0,0,0],[9E+09,9E+09,9E+09,9E+09,9E+09,9E+09]];
    CONST robtarget Target_2340:=[[108.478856861,140.459552219,0],[0.882142515,0,0,-0.470982573],[0,0,0,0],[9E+09,9E+09,9E+09,9E+09,9E+09,9E+09]];
    CONST robtarget Target_2350:=[[106.60526948,142.674933361,0],[0.882142515,0,0,-0.470982573],[0,0,0,0],[9E+09,9E+09,9E+09,9E+09,9E+09,9E+09]];
    CONST robtarget Target_2360:=[[109.768501207,141.609028207,0],[0.882142515,0,0,-0.470982573],[0,0,0,0],[9E+09,9E+09,9E+09,9E+09,9E+09,9E+09]];
    CONST robtarget Target_2370:=[[112.752717891,141.326992858,0],[0.882142515,0,0,-0.470982573],[0,0,0,0],[9E+09,9E+09,9E+09,9E+09,9E+09,9E+09]];
    CONST robtarget Target_2380:=[[115.631258945,142.163111606,0],[0.882142515,0,0,-0.470982573],[0,0,0,0],[9E+09,9E+09,9E+09,9E+09,9E+09,9E+09]];
    CONST robtarget Target_2390:=[[118,144,0],[0.882142515,0,0,-0.470982573],[0,0,0,0],[9E+09,9E+09,9E+09,9E+09,9E+09,9E+09]];
    CONST robtarget Target_2400:=[[115.336324555,142.849749419,0],[0.882142515,0,0,-0.470982573],[0,0,0,0],[9E+09,9E+09,9E+09,9E+09,9E+09,9E+09]];
    CONST robtarget Target_2410:=[[112.437578714,142.725186884,0],[0.882142515,0,0,-0.470982573],[0,0,0,0],[9E+09,9E+09,9E+09,9E+09,9E+09,9E+09]];
    CONST robtarget Target_2420:=[[109.685049159,143.642696736,0],[0.882142515,0,0,-0.470982573],[0,0,0,0],[9E+09,9E+09,9E+09,9E+09,9E+09,9E+09]];
    CONST robtarget Target_2430:=[[107.440790007,145.481594268,0],[0.882142515,0,0,-0.470982573],[0,0,0,0],[9E+09,9E+09,9E+09,9E+09,9E+09,9E+09]];
    CONST robtarget Target_2440:=[[106,148,0],[0.882142515,0,0,-0.470982573],[0,0,0,0],[9E+09,9E+09,9E+09,9E+09,9E+09,9E+09]];
    CONST robtarget Target_2450:=[[108.368741055,146.163111606,0],[0.882142515,0,0,-0.470982573],[0,0,0,0],[9E+09,9E+09,9E+09,9E+09,9E+09,9E+09]];
    CONST robtarget Target_2460:=[[111.247282109,145.326992858,0],[0.882142515,0,0,-0.470982573],[0,0,0,0],[9E+09,9E+09,9E+09,9E+09,9E+09,9E+09]];
    CONST robtarget Target_2470:=[[114.231498793,145.609028207,0],[0.882142515,0,0,-0.470982573],[0,0,0,0],[9E+09,9E+09,9E+09,9E+09,9E+09,9E+09]];
    CONST robtarget Target_2480:=[[116.902430719,146.969622123,0],[0.882142515,0,0,-0.470982573],[0,0,0,0],[9E+09,9E+09,9E+09,9E+09,9E+09,9E+09]];
    CONST robtarget Target_2490:=[[113.892645843,146.654955892,0],[0.882142515,0,0,-0.470982573],[0,0,0,0],[9E+09,9E+09,9E+09,9E+09,9E+09,9E+09]];
    CONST robtarget Target_2500:=[[111.01937121,147.058113631,0],[0.882142515,0,0,-0.470982573],[0,0,0,0],[9E+09,9E+09,9E+09,9E+09,9E+09,9E+09]];
    CONST robtarget Target_2510:=[[108.478856861,148.459552219,0],[0.882142515,0,0,-0.470982573],[0,0,0,0],[9E+09,9E+09,9E+09,9E+09,9E+09,9E+09]];
    CONST robtarget Target_2520:=[[106.60526948,150.674933361,0],[0.882142515,0,0,-0.470982573],[0,0,0,0],[9E+09,9E+09,9E+09,9E+09,9E+09,9E+09]];
    CONST robtarget Target_2530:=[[109.768501207,149.609028207,0],[0.882142515,0,0,-0.470982573],[0,0,0,0],[9E+09,9E+09,9E+09,9E+09,9E+09,9E+09]];
    CONST robtarget Target_2540:=[[112.752717891,149.326992858,0],[0.882142515,0,0,-0.470982573],[0,0,0,0],[9E+09,9E+09,9E+09,9E+09,9E+09,9E+09]];
    CONST robtarget Target_2550:=[[115.631258945,150.163111606,0],[0.882142515,0,0,-0.470982573],[0,0,0,0],[9E+09,9E+09,9E+09,9E+09,9E+09,9E+09]];
    CONST robtarget Target_2560:=[[118,152,0],[0.882142515,0,0,-0.470982573],[0,0,0,0],[9E+09,9E+09,9E+09,9E+09,9E+09,9E+09]];
    CONST robtarget Target_2570:=[[115.336324555,150.849749419,0],[0.882142515,0,0,-0.470982573],[0,0,0,0],[9E+09,9E+09,9E+09,9E+09,9E+09,9E+09]];
    CONST robtarget Target_2580:=[[112.437578714,150.725186884,0],[0.882142515,0,0,-0.470982573],[0,0,0,0],[9E+09,9E+09,9E+09,9E+09,9E+09,9E+09]];
    CONST robtarget Target_2590:=[[109.685049159,151.642696736,0],[0.882142515,0,0,-0.470982573],[0,0,0,0],[9E+09,9E+09,9E+09,9E+09,9E+09,9E+09]];
    CONST robtarget Target_2600:=[[107.440790007,153.481594268,0],[0.882142515,0,0,-0.470982573],[0,0,0,0],[9E+09,9E+09,9E+09,9E+09,9E+09,9E+09]];
    CONST robtarget Target_2610:=[[106,156,0],[0.882142515,0,0,-0.470982573],[0,0,0,0],[9E+09,9E+09,9E+09,9E+09,9E+09,9E+09]];
    CONST robtarget Target_2620:=[[108.368741055,154.163111606,0],[0.882142515,0,0,-0.470982573],[0,0,0,0],[9E+09,9E+09,9E+09,9E+09,9E+09,9E+09]];
    CONST robtarget Target_2630:=[[111.247282109,153.326992858,0],[0.882142515,0,0,-0.470982573],[0,0,0,0],[9E+09,9E+09,9E+09,9E+09,9E+09,9E+09]];
    CONST robtarget Target_2640:=[[114.231498793,153.609028207,0],[0.882142515,0,0,-0.470982573],[0,0,0,0],[9E+09,9E+09,9E+09,9E+09,9E+09,9E+09]];
    CONST robtarget Target_2650:=[[116.902430719,154.969622123,0],[0.882142515,0,0,-0.470982573],[0,0,0,0],[9E+09,9E+09,9E+09,9E+09,9E+09,9E+09]];
    CONST robtarget Target_2660:=[[113.892645843,154.654955892,0],[0.882142515,0,0,-0.470982573],[0,0,0,0],[9E+09,9E+09,9E+09,9E+09,9E+09,9E+09]];
    CONST robtarget Target_2670:=[[111.01937121,155.058113631,0],[0.882142515,0,0,-0.470982573],[0,0,0,0],[9E+09,9E+09,9E+09,9E+09,9E+09,9E+09]];
    CONST robtarget Target_2680:=[[108.478856861,156.459552219,0],[0.882142515,0,0,-0.470982573],[0,0,0,0],[9E+09,9E+09,9E+09,9E+09,9E+09,9E+09]];
    CONST robtarget Target_2690:=[[106.60526948,158.674933361,0],[0.882142515,0,0,-0.470982573],[0,0,0,0],[9E+09,9E+09,9E+09,9E+09,9E+09,9E+09]];
    CONST robtarget Target_2700:=[[109.768501207,157.609028207,0],[0.882142515,0,0,-0.470982573],[0,0,0,0],[9E+09,9E+09,9E+09,9E+09,9E+09,9E+09]];
    CONST robtarget Target_2710:=[[112.752717891,157.326992858,0],[0.882142515,0,0,-0.470982573],[0,0,0,0],[9E+09,9E+09,9E+09,9E+09,9E+09,9E+09]];
    CONST robtarget Target_2720:=[[115.631258945,158.163111606,0],[0.882142515,0,0,-0.470982573],[0,0,0,0],[9E+09,9E+09,9E+09,9E+09,9E+09,9E+09]];
    CONST robtarget Target_2730:=[[118,160,0],[0.882142515,0,0,-0.470982573],[0,0,0,0],[9E+09,9E+09,9E+09,9E+09,9E+09,9E+09]];
    CONST robtarget Target_2740:=[[115.336324555,158.849749419,0],[0.882142515,0,0,-0.470982573],[0,0,0,0],[9E+09,9E+09,9E+09,9E+09,9E+09,9E+09]];
    CONST robtarget Target_2750:=[[112.437578714,158.725186884,0],[0.882142515,0,0,-0.470982573],[0,0,0,0],[9E+09,9E+09,9E+09,9E+09,9E+09,9E+09]];
    CONST robtarget Target_2760:=[[109.685049159,159.642696736,0],[0.882142515,0,0,-0.470982573],[0,0,0,0],[9E+09,9E+09,9E+09,9E+09,9E+09,9E+09]];
    CONST robtarget Target_2770:=[[107.440790007,161.481594268,0],[0.882142515,0,0,-0.470982573],[0,0,0,0],[9E+09,9E+09,9E+09,9E+09,9E+09,9E+09]];
    CONST robtarget Target_2780:=[[106,164,0],[0.882142515,0,0,-0.470982573],[0,0,0,0],[9E+09,9E+09,9E+09,9E+09,9E+09,9E+09]];
    CONST robtarget Target_2790:=[[108.368741055,162.163111606,0],[0.882142515,0,0,-0.470982573],[0,0,0,0],[9E+09,9E+09,9E+09,9E+09,9E+09,9E+09]];
    CONST robtarget Target_2800:=[[111.247282109,161.326992858,0],[0.882142515,0,0,-0.470982573],[0,0,0,0],[9E+09,9E+09,9E+09,9E+09,9E+09,9E+09]];
    CONST robtarget Target_2810:=[[114.231498793,161.609028207,0],[0.882142515,0,0,-0.470982573],[0,0,0,0],[9E+09,9E+09,9E+09,9E+09,9E+09,9E+09]];
    CONST robtarget Target_2820:=[[116.902430719,162.969622123,0],[0.882142515,0,0,-0.470982573],[0,0,0,0],[9E+09,9E+09,9E+09,9E+09,9E+09,9E+09]];
    CONST robtarget Target_2830:=[[113.892645843,162.654955892,0],[0.882142515,0,0,-0.470982573],[0,0,0,0],[9E+09,9E+09,9E+09,9E+09,9E+09,9E+09]];
    CONST robtarget Target_2840:=[[111.01937121,163.058113631,0],[0.882142515,0,0,-0.470982573],[0,0,0,0],[9E+09,9E+09,9E+09,9E+09,9E+09,9E+09]];
    CONST robtarget Target_2850:=[[108.478856861,164.459552219,0],[0.882142515,0,0,-0.470982573],[0,0,0,0],[9E+09,9E+09,9E+09,9E+09,9E+09,9E+09]];
    CONST robtarget Target_2860:=[[106.60526948,166.674933361,0],[0.882142515,0,0,-0.470982573],[0,0,0,0],[9E+09,9E+09,9E+09,9E+09,9E+09,9E+09]];
    CONST robtarget Target_2870:=[[109.768501207,165.609028207,0],[0.882142515,0,0,-0.470982573],[0,0,0,0],[9E+09,9E+09,9E+09,9E+09,9E+09,9E+09]];
    CONST robtarget Target_2880:=[[112.752717891,165.326992858,0],[0.882142515,0,0,-0.470982573],[0,0,0,0],[9E+09,9E+09,9E+09,9E+09,9E+09,9E+09]];
    CONST robtarget Target_2890:=[[115.631258945,166.163111606,0],[0.882142515,0,0,-0.470982573],[0,0,0,0],[9E+09,9E+09,9E+09,9E+09,9E+09,9E+09]];
    CONST robtarget Target_2900:=[[118,168,0],[0.882142515,0,0,-0.470982573],[0,0,0,0],[9E+09,9E+09,9E+09,9E+09,9E+09,9E+09]];
    CONST robtarget Target_2910:=[[115.336324555,166.849749419,0],[0.882142515,0,0,-0.470982573],[0,0,0,0],[9E+09,9E+09,9E+09,9E+09,9E+09,9E+09]];
    CONST robtarget Target_2920:=[[112.437578714,166.725186884,0],[0.882142515,0,0,-0.470982573],[0,0,0,0],[9E+09,9E+09,9E+09,9E+09,9E+09,9E+09]];
    CONST robtarget Target_2930:=[[109.685049159,167.642696736,0],[0.882142515,0,0,-0.470982573],[0,0,0,0],[9E+09,9E+09,9E+09,9E+09,9E+09,9E+09]];
    CONST robtarget Target_2940:=[[107.440790007,169.481594268,0],[0.882142515,0,0,-0.470982573],[0,0,0,0],[9E+09,9E+09,9E+09,9E+09,9E+09,9E+09]];
    CONST robtarget Target_2950:=[[106,172,0],[0.882142515,0,0,-0.470982573],[0,0,0,0],[9E+09,9E+09,9E+09,9E+09,9E+09,9E+09]];
    CONST robtarget Target_2960:=[[108.368741055,170.163111606,0],[0.882142515,0,0,-0.470982573],[0,0,0,0],[9E+09,9E+09,9E+09,9E+09,9E+09,9E+09]];
    CONST robtarget Target_2970:=[[111.247282109,169.326992858,0],[0.882142515,0,0,-0.470982573],[0,0,0,0],[9E+09,9E+09,9E+09,9E+09,9E+09,9E+09]];
    CONST robtarget Target_2980:=[[114.231498793,169.609028207,0],[0.882142515,0,0,-0.470982573],[0,0,0,0],[9E+09,9E+09,9E+09,9E+09,9E+09,9E+09]];
    CONST robtarget Target_2990:=[[116.902430719,170.969622123,0],[0.882142515,0,0,-0.470982573],[0,0,0,0],[9E+09,9E+09,9E+09,9E+09,9E+09,9E+09]];
    CONST robtarget Target_3000:=[[113.892645843,170.654955892,0],[0.882142515,0,0,-0.470982573],[0,0,0,0],[9E+09,9E+09,9E+09,9E+09,9E+09,9E+09]];
    CONST robtarget Target_3010:=[[111.01937121,171.058113631,0],[0.882142515,0,0,-0.470982573],[0,0,0,0],[9E+09,9E+09,9E+09,9E+09,9E+09,9E+09]];
    CONST robtarget Target_3020:=[[108.478856861,172.459552219,0],[0.882142515,0,0,-0.470982573],[0,0,0,0],[9E+09,9E+09,9E+09,9E+09,9E+09,9E+09]];
    CONST robtarget Target_3030:=[[106.60526948,174.674933361,0],[0.882142515,0,0,-0.470982573],[0,0,0,0],[9E+09,9E+09,9E+09,9E+09,9E+09,9E+09]];
    CONST robtarget Target_3040:=[[109.768501207,173.609028207,0],[0.882142515,0,0,-0.470982573],[0,0,0,0],[9E+09,9E+09,9E+09,9E+09,9E+09,9E+09]];
    CONST robtarget Target_3050:=[[112.752717891,173.326992858,0],[0.882142515,0,0,-0.470982573],[0,0,0,0],[9E+09,9E+09,9E+09,9E+09,9E+09,9E+09]];
    CONST robtarget Target_3070:=[[118,176,0],[0.882142515,0,0,-0.470982573],[0,0,0,0],[9E+09,9E+09,9E+09,9E+09,9E+09,9E+09]];
    CONST robtarget Target_3080:=[[115.336324555,174.849749419,0],[0.882142515,0,0,-0.470982573],[0,0,0,0],[9E+09,9E+09,9E+09,9E+09,9E+09,9E+09]];
    CONST robtarget Target_3090:=[[112.437578714,174.725186884,0],[0.882142515,0,0,-0.470982573],[0,0,0,0],[9E+09,9E+09,9E+09,9E+09,9E+09,9E+09]];
    CONST robtarget Target_3100:=[[109.685049159,175.642696736,0],[0.882142515,0,0,-0.470982573],[0,0,0,0],[9E+09,9E+09,9E+09,9E+09,9E+09,9E+09]];
    CONST robtarget Target_3110:=[[107.440790007,177.481594268,0],[0.882142515,0,0,-0.470982573],[0,0,0,0],[9E+09,9E+09,9E+09,9E+09,9E+09,9E+09]];
    CONST robtarget Target_3120:=[[106,180,0],[0.882142515,0,0,-0.470982573],[0,0,0,0],[9E+09,9E+09,9E+09,9E+09,9E+09,9E+09]];
    CONST robtarget Target_3130:=[[108.368741055,178.163111606,0],[0.882142515,0,0,-0.470982573],[0,0,0,0],[9E+09,9E+09,9E+09,9E+09,9E+09,9E+09]];
    CONST robtarget Target_3140:=[[111.247282109,177.326992858,0],[0.882142515,0,0,-0.470982573],[0,0,0,0],[9E+09,9E+09,9E+09,9E+09,9E+09,9E+09]];
    CONST robtarget Target_3150:=[[114.231498793,177.609028207,0],[0.882142515,0,0,-0.470982573],[0,0,0,0],[9E+09,9E+09,9E+09,9E+09,9E+09,9E+09]];
    CONST robtarget Target_3160:=[[116.902430719,178.969622123,0],[0.882142515,0,0,-0.470982573],[0,0,0,0],[9E+09,9E+09,9E+09,9E+09,9E+09,9E+09]];
    CONST robtarget Target_3170:=[[118,180,0],[0.882142515,0,0,-0.470982573],[0,0,0,0],[9E+09,9E+09,9E+09,9E+09,9E+09,9E+09]];
    CONST robtarget Target_3060:=[[115.631258945,174.163111606,0],[0.882142515,0,0,-0.470982573],[0,0,0,0],[9E+09,9E+09,9E+09,9E+09,9E+09,9E+09]];
    CONST robtarget Target_3180:=[[76.943222938,151.35527551,0],[0.882142515,0,0,-0.470982573],[0,0,0,0],[9E+09,9E+09,9E+09,9E+09,9E+09,9E+09]];
    CONST robtarget Target_3190:=[[65.513222871,151.35527551,0],[0.882142515,0,0,-0.470982573],[0,0,0,0],[9E+09,9E+09,9E+09,9E+09,9E+09,9E+09]];
    CONST robtarget Target_3200:=[[65.513222871,148.752495916,0],[0.882142515,0,0,-0.470982573],[0,0,0,0],[9E+09,9E+09,9E+09,9E+09,9E+09,9E+09]];
    CONST robtarget Target_3210:=[[65.573429517,147.314483347,0],[0.882142515,0,0,-0.470982573],[0,0,0,0],[9E+09,9E+09,9E+09,9E+09,9E+09,9E+09]];
    CONST robtarget Target_3220:=[[65.754049453,146.223816809,0],[0.882142515,0,0,-0.470982573],[0,0,0,0],[9E+09,9E+09,9E+09,9E+09,9E+09,9E+09]];
    CONST robtarget Target_3230:=[[66.420953833,144.658444028,0],[0.882142515,0,0,-0.470982573],[0,0,0,0],[9E+09,9E+09,9E+09,9E+09,9E+09,9E+09]];
    CONST robtarget Target_3240:=[[67.271951609,143.68008604,0],[0.882142515,0,0,-0.470982573],[0,0,0,0],[9E+09,9E+09,9E+09,9E+09,9E+09,9E+09]];
    CONST robtarget Target_3250:=[[68.361460327,142.949501554,0],[0.882142515,0,0,-0.470982573],[0,0,0,0],[9E+09,9E+09,9E+09,9E+09,9E+09,9E+09]];
    CONST robtarget Target_3260:=[[69.684848706,142.494478254,0],[0.882142515,0,0,-0.470982573],[0,0,0,0],[9E+09,9E+09,9E+09,9E+09,9E+09,9E+09]];
    CONST robtarget Target_3270:=[[71.237485465,142.34280382,0],[0.882142515,0,0,-0.470982573],[0,0,0,0],[9E+09,9E+09,9E+09,9E+09,9E+09,9E+09]];
    CONST robtarget Target_3280:=[[72.726442119,142.501425174,0],[0.882142515,0,0,-0.470982573],[0,0,0,0],[9E+09,9E+09,9E+09,9E+09,9E+09,9E+09]];
    CONST robtarget Target_3290:=[[74.062566519,142.977289237,0],[0.882142515,0,0,-0.470982573],[0,0,0,0],[9E+09,9E+09,9E+09,9E+09,9E+09,9E+09]];
    CONST robtarget Target_3300:=[[75.18333638,143.719451924,0],[0.882142515,0,0,-0.470982573],[0,0,0,0],[9E+09,9E+09,9E+09,9E+09,9E+09,9E+09]];
    CONST robtarget Target_3310:=[[76.026229416,144.67696915,0],[0.882142515,0,0,-0.470982573],[0,0,0,0],[9E+09,9E+09,9E+09,9E+09,9E+09,9E+09]];
    CONST robtarget Target_3320:=[[76.757971721,146.441486988,0],[0.882142515,0,0,-0.470982573],[0,0,0,0],[9E+09,9E+09,9E+09,9E+09,9E+09,9E+09]];
    CONST robtarget Target_3330:=[[76.896910134,147.45921086,0],[0.882142515,0,0,-0.470982573],[0,0,0,0],[9E+09,9E+09,9E+09,9E+09,9E+09,9E+09]];
    CONST robtarget Target_3340:=[[76.943222938,148.724708233,0],[0.882142515,0,0,-0.470982573],[0,0,0,0],[9E+09,9E+09,9E+09,9E+09,9E+09,9E+09]];
    CONST robtarget Target_3350:=[[76.943222938,151.35527551,0],[0.882142515,0,0,-0.470982573],[0,0,0,0],[9E+09,9E+09,9E+09,9E+09,9E+09,9E+09]];
    CONST robtarget Target_3360:=[[66.828506509,149.836215533,0],[0.882142515,0,0,-0.470982573],[0,0,0,0],[9E+09,9E+09,9E+09,9E+09,9E+09,9E+09]];
    CONST robtarget Target_3370:=[[66.828506509,148.678395429,0],[0.882142515,0,0,-0.470982573],[0,0,0,0],[9E+09,9E+09,9E+09,9E+09,9E+09,9E+09]];
    CONST robtarget Target_3380:=[[66.990601324,146.960190395,0],[0.882142515,0,0,-0.470982573],[0,0,0,0],[9E+09,9E+09,9E+09,9E+09,9E+09,9E+09]];
    CONST robtarget Target_3390:=[[67.513936011,145.658800598,0],[0.882142515,0,0,-0.470982573],[0,0,0,0],[9E+09,9E+09,9E+09,9E+09,9E+09,9E+09]];
    CONST robtarget Target_3400:=[[68.972789342,144.362042081,0],[0.882142515,0,0,-0.470982573],[0,0,0,0],[9E+09,9E+09,9E+09,9E+09,9E+09,9E+09]];
    CONST robtarget Target_3410:=[[69.999775774,144.035536812,0],[0.882142515,0,0,-0.470982573],[0,0,0,0],[9E+09,9E+09,9E+09,9E+09,9E+09,9E+09]];
    CONST robtarget Target_3420:=[[71.218960344,143.926701722,0],[0.882142515,0,0,-0.470982573],[0,0,0,0],[9E+09,9E+09,9E+09,9E+09,9E+09,9E+09]];
    CONST robtarget Target_3430:=[[72.441618374,144.026274251,0],[0.882142515,0,0,-0.470982573],[0,0,0,0],[9E+09,9E+09,9E+09,9E+09,9E+09,9E+09]];
    CONST robtarget Target_3440:=[[73.441974943,144.324991838,0],[0.882142515,0,0,-0.470982573],[0,0,0,0],[9E+09,9E+09,9E+09,9E+09,9E+09,9E+09]];
    CONST robtarget Target_3450:=[[74.868409312,145.519862185,0],[0.882142515,0,0,-0.470982573],[0,0,0,0],[9E+09,9E+09,9E+09,9E+09,9E+09,9E+09]];
    CONST robtarget Target_3460:=[[75.465844485,146.90461503,0],[0.882142515,0,0,-0.470982573],[0,0,0,0],[9E+09,9E+09,9E+09,9E+09,9E+09,9E+09]];
    CONST robtarget Target_3470:=[[75.6279393,148.678395429,0],[0.882142515,0,0,-0.470982573],[0,0,0,0],[9E+09,9E+09,9E+09,9E+09,9E+09,9E+09]];
    CONST robtarget Target_3480:=[[75.6279393,149.836215533,0],[0.882142515,0,0,-0.470982573],[0,0,0,0],[9E+09,9E+09,9E+09,9E+09,9E+09,9E+09]];
    CONST robtarget Target_3490:=[[66.828506509,149.836215533,0],[0.882142515,0,0,-0.470982573],[0,0,0,0],[9E+09,9E+09,9E+09,9E+09,9E+09,9E+09]];
    CONST robtarget Target_3500:=[[72.451,138.934,0],[0.882142515,0,0,-0.470982573],[0,0,0,0],[9E+09,9E+09,9E+09,9E+09,9E+09,9E+09]];
    CONST robtarget Target_3510:=[[67.069,137.174,0],[0.882142515,0,0,-0.470982573],[0,0,0,0],[9E+09,9E+09,9E+09,9E+09,9E+09,9E+09]];
    CONST robtarget Target_3520:=[[72.451,135.405,0],[0.882142515,0,0,-0.470982573],[0,0,0,0],[9E+09,9E+09,9E+09,9E+09,9E+09,9E+09]];
    CONST robtarget Target_3530:=[[76.943222938,141.925988583,0],[0.882142515,0,0,-0.470982573],[0,0,0,0],[9E+09,9E+09,9E+09,9E+09,9E+09,9E+09]];
    CONST robtarget Target_3540:=[[65.513222871,138.072763276,0],[0.882142515,0,0,-0.470982573],[0,0,0,0],[9E+09,9E+09,9E+09,9E+09,9E+09,9E+09]];
    CONST robtarget Target_3550:=[[65.513222871,136.201725988,0],[0.882142515,0,0,-0.470982573],[0,0,0,0],[9E+09,9E+09,9E+09,9E+09,9E+09,9E+09]];
    CONST robtarget Target_3560:=[[76.943222938,132.348500682,0],[0.882142515,0,0,-0.470982573],[0,0,0,0],[9E+09,9E+09,9E+09,9E+09,9E+09,9E+09]];
    CONST robtarget Target_3570:=[[76.943222938,133.950923706,0],[0.882142515,0,0,-0.470982573],[0,0,0,0],[9E+09,9E+09,9E+09,9E+09,9E+09,9E+09]];
    CONST robtarget Target_3580:=[[73.747639451,134.988330519,0],[0.882142515,0,0,-0.470982573],[0,0,0,0],[9E+09,9E+09,9E+09,9E+09,9E+09,9E+09]];
    CONST robtarget Target_3590:=[[73.747639451,139.350996671,0],[0.882142515,0,0,-0.470982573],[0,0,0,0],[9E+09,9E+09,9E+09,9E+09,9E+09,9E+09]];
    CONST robtarget Target_3600:=[[76.943222938,140.388403484,0],[0.882142515,0,0,-0.470982573],[0,0,0,0],[9E+09,9E+09,9E+09,9E+09,9E+09,9E+09]];
    CONST robtarget Target_3610:=[[76.943222938,141.925988583,0],[0.882142515,0,0,-0.470982573],[0,0,0,0],[9E+09,9E+09,9E+09,9E+09,9E+09,9E+09]];
    CONST robtarget Target_3620:=[[65.513222871,130.857228388,0],[0.882142515,0,0,-0.470982573],[0,0,0,0],[9E+09,9E+09,9E+09,9E+09,9E+09,9E+09]];
    CONST robtarget Target_3630:=[[65.513222871,132.487439095,0],[0.882142515,0,0,-0.470982573],[0,0,0,0],[9E+09,9E+09,9E+09,9E+09,9E+09,9E+09]];
    CONST robtarget Target_3640:=[[76.943222938,128.550850741,0],[0.882142515,0,0,-0.470982573],[0,0,0,0],[9E+09,9E+09,9E+09,9E+09,9E+09,9E+09]];
    CONST robtarget Target_3650:=[[76.943222938,126.911377474,0],[0.882142515,0,0,-0.470982573],[0,0,0,0],[9E+09,9E+09,9E+09,9E+09,9E+09,9E+09]];
    CONST robtarget Target_3660:=[[65.513222871,122.97478912,0],[0.882142515,0,0,-0.470982573],[0,0,0,0],[9E+09,9E+09,9E+09,9E+09,9E+09,9E+09]];
    CONST robtarget Target_3670:=[[65.513222871,124.521636779,0],[0.882142515,0,0,-0.470982573],[0,0,0,0],[9E+09,9E+09,9E+09,9E+09,9E+09,9E+09]];
    CONST robtarget Target_3680:=[[75.007347724,127.689432584,0],[0.882142515,0,0,-0.470982573],[0,0,0,0],[9E+09,9E+09,9E+09,9E+09,9E+09,9E+09]];
    CONST robtarget Target_3690:=[[65.513222871,130.857228388,0],[0.882142515,0,0,-0.470982573],[0,0,0,0],[9E+09,9E+09,9E+09,9E+09,9E+09,9E+09]];
    CONST robtarget Target_3820:=[[65.513,122.326,0],[0.882142515,0,0,-0.470982573],[0,0,0,0],[9E+09,9E+09,9E+09,9E+09,9E+09,9E+09]];
    CONST robtarget Target_3810:=[[65.513,117.899,0],[0.882142515,0,0,-0.470982573],[0,0,0,0],[9E+09,9E+09,9E+09,9E+09,9E+09,9E+09]];
    CONST robtarget Target_3800:=[[66.68,117.899,0],[0.882142515,0,0,-0.470982573],[0,0,0,0],[9E+09,9E+09,9E+09,9E+09,9E+09,9E+09]];
    CONST robtarget Target_3790:=[[66.68,119.353,0],[0.882142515,0,0,-0.470982573],[0,0,0,0],[9E+09,9E+09,9E+09,9E+09,9E+09,9E+09]];
    CONST robtarget Target_3780:=[[75.776,119.353,0],[0.882142515,0,0,-0.470982573],[0,0,0,0],[9E+09,9E+09,9E+09,9E+09,9E+09,9E+09]];
    CONST robtarget Target_3770:=[[75.776,117.899,0],[0.882142515,0,0,-0.470982573],[0,0,0,0],[9E+09,9E+09,9E+09,9E+09,9E+09,9E+09]];
    CONST robtarget Target_3760:=[[76.943,117.899,0],[0.882142515,0,0,-0.470982573],[0,0,0,0],[9E+09,9E+09,9E+09,9E+09,9E+09,9E+09]];
    CONST robtarget Target_3750:=[[76.943,122.326,0],[0.882142515,0,0,-0.470982573],[0,0,0,0],[9E+09,9E+09,9E+09,9E+09,9E+09,9E+09]];
    CONST robtarget Target_3740:=[[75.776,122.326,0],[0.882142515,0,0,-0.470982573],[0,0,0,0],[9E+09,9E+09,9E+09,9E+09,9E+09,9E+09]];
    CONST robtarget Target_3730:=[[75.776,120.872,0],[0.882142515,0,0,-0.470982573],[0,0,0,0],[9E+09,9E+09,9E+09,9E+09,9E+09,9E+09]];
    CONST robtarget Target_3720:=[[66.68,120.872,0],[0.882142515,0,0,-0.470982573],[0,0,0,0],[9E+09,9E+09,9E+09,9E+09,9E+09,9E+09]];
    CONST robtarget Target_3710:=[[66.68,122.326,0],[0.882142515,0,0,-0.470982573],[0,0,0,0],[9E+09,9E+09,9E+09,9E+09,9E+09,9E+09]];
    CONST robtarget Target_3700:=[[65.513,122.326,0],[0.882142515,0,0,-0.470982573],[0,0,0,0],[9E+09,9E+09,9E+09,9E+09,9E+09,9E+09]];
    CONST robtarget Target_3830:=[[65.513222871,116.018605935,0],[0.882142515,0,0,-0.470982573],[0,0,0,0],[9E+09,9E+09,9E+09,9E+09,9E+09,9E+09]];
    CONST robtarget Target_3840:=[[65.513222871,113.415826341,0],[0.882142515,0,0,-0.470982573],[0,0,0,0],[9E+09,9E+09,9E+09,9E+09,9E+09,9E+09]];
    CONST robtarget Target_3850:=[[65.516985787,113.023759509,0],[0.882142515,0,0,-0.470982573],[0,0,0,0],[9E+09,9E+09,9E+09,9E+09,9E+09,9E+09]];
    CONST robtarget Target_3860:=[[65.528274533,112.653401803,0],[0.882142515,0,0,-0.470982573],[0,0,0,0],[9E+09,9E+09,9E+09,9E+09,9E+09,9E+09]];
    CONST robtarget Target_3870:=[[65.547089109,112.304753224,0],[0.882142515,0,0,-0.470982573],[0,0,0,0],[9E+09,9E+09,9E+09,9E+09,9E+09,9E+09]];
    CONST robtarget Target_3880:=[[65.573429517,111.977813772,0],[0.882142515,0,0,-0.470982573],[0,0,0,0],[9E+09,9E+09,9E+09,9E+09,9E+09,9E+09]];
    CONST robtarget Target_3890:=[[65.607295755,111.672583447,0],[0.882142515,0,0,-0.470982573],[0,0,0,0],[9E+09,9E+09,9E+09,9E+09,9E+09,9E+09]];
    CONST robtarget Target_3900:=[[65.648687823,111.389062249,0],[0.882142515,0,0,-0.470982573],[0,0,0,0],[9E+09,9E+09,9E+09,9E+09,9E+09,9E+09]];
    CONST robtarget Target_3910:=[[65.697605723,111.127250178,0],[0.882142515,0,0,-0.470982573],[0,0,0,0],[9E+09,9E+09,9E+09,9E+09,9E+09,9E+09]];
    CONST robtarget Target_3920:=[[65.754049453,110.887147234,0],[0.882142515,0,0,-0.470982573],[0,0,0,0],[9E+09,9E+09,9E+09,9E+09,9E+09,9E+09]];
    CONST robtarget Target_3930:=[[65.886040945,110.445438865,0],[0.882142515,0,0,-0.470982573],[0,0,0,0],[9E+09,9E+09,9E+09,9E+09,9E+09,9E+09]];
    CONST robtarget Target_3940:=[[66.041188839,110.037307278,0],[0.882142515,0,0,-0.470982573],[0,0,0,0],[9E+09,9E+09,9E+09,9E+09,9E+09,9E+09]];
    CONST robtarget Target_3950:=[[66.219493135,109.662752474,0],[0.882142515,0,0,-0.470982573],[0,0,0,0],[9E+09,9E+09,9E+09,9E+09,9E+09,9E+09]];
    CONST robtarget Target_3960:=[[66.420953833,109.321774454,0],[0.882142515,0,0,-0.470982573],[0,0,0,0],[9E+09,9E+09,9E+09,9E+09,9E+09,9E+09]];
    CONST robtarget Target_3970:=[[66.611342876,109.053956191,0],[0.882142515,0,0,-0.470982573],[0,0,0,0],[9E+09,9E+09,9E+09,9E+09,9E+09,9E+09]];
    CONST robtarget Target_3980:=[[66.816638853,108.801623772,0],[0.882142515,0,0,-0.470982573],[0,0,0,0],[9E+09,9E+09,9E+09,9E+09,9E+09,9E+09]];
    CONST robtarget Target_3990:=[[67.036841764,108.564777197,0],[0.882142515,0,0,-0.470982573],[0,0,0,0],[9E+09,9E+09,9E+09,9E+09,9E+09,9E+09]];
    CONST robtarget Target_4000:=[[67.271951609,108.343416466,0],[0.882142515,0,0,-0.470982573],[0,0,0,0],[9E+09,9E+09,9E+09,9E+09,9E+09,9E+09]];
    CONST robtarget Target_4010:=[[67.521968388,108.137541579,0],[0.882142515,0,0,-0.470982573],[0,0,0,0],[9E+09,9E+09,9E+09,9E+09,9E+09,9E+09]];
    CONST robtarget Target_4020:=[[67.786892101,107.947152535,0],[0.882142515,0,0,-0.470982573],[0,0,0,0],[9E+09,9E+09,9E+09,9E+09,9E+09,9E+09]];
    CONST robtarget Target_4030:=[[68.066722747,107.772249336,0],[0.882142515,0,0,-0.470982573],[0,0,0,0],[9E+09,9E+09,9E+09,9E+09,9E+09,9E+09]];
    CONST robtarget Target_4040:=[[68.361460327,107.61283198,0],[0.882142515,0,0,-0.470982573],[0,0,0,0],[9E+09,9E+09,9E+09,9E+09,9E+09,9E+09]];
    CONST robtarget Target_4050:=[[68.670815386,107.470637199,0],[0.882142515,0,0,-0.470982573],[0,0,0,0],[9E+09,9E+09,9E+09,9E+09,9E+09,9E+09]];
    CONST robtarget Target_4060:=[[68.994498469,107.347401721,0],[0.882142515,0,0,-0.470982573],[0,0,0,0],[9E+09,9E+09,9E+09,9E+09,9E+09,9E+09]];
    CONST robtarget Target_4070:=[[69.332509576,107.243125548,0],[0.882142515,0,0,-0.470982573],[0,0,0,0],[9E+09,9E+09,9E+09,9E+09,9E+09,9E+09]];
    CONST robtarget Target_4080:=[[69.684848706,107.157808679,0],[0.882142515,0,0,-0.470982573],[0,0,0,0],[9E+09,9E+09,9E+09,9E+09,9E+09,9E+09]];
    CONST robtarget Target_4090:=[[70.05151586,107.091451115,0],[0.882142515,0,0,-0.470982573],[0,0,0,0],[9E+09,9E+09,9E+09,9E+09,9E+09,9E+09]];
    CONST robtarget Target_4100:=[[70.432511038,107.044052854,0],[0.882142515,0,0,-0.470982573],[0,0,0,0],[9E+09,9E+09,9E+09,9E+09,9E+09,9E+09]];
    CONST robtarget Target_4110:=[[70.82783424,107.015613898,0],[0.882142515,0,0,-0.470982573],[0,0,0,0],[9E+09,9E+09,9E+09,9E+09,9E+09,9E+09]];
    CONST robtarget Target_4120:=[[71.237485465,107.006134246,0],[0.882142515,0,0,-0.470982573],[0,0,0,0],[9E+09,9E+09,9E+09,9E+09,9E+09,9E+09]];
    CONST robtarget Target_4130:=[[71.624052653,107.01604808,0],[0.882142515,0,0,-0.470982573],[0,0,0,0],[9E+09,9E+09,9E+09,9E+09,9E+09,9E+09]];
    CONST robtarget Target_4140:=[[72.001067824,107.045789584,0],[0.882142515,0,0,-0.470982573],[0,0,0,0],[9E+09,9E+09,9E+09,9E+09,9E+09,9E+09]];
    CONST robtarget Target_4150:=[[72.36853098,107.095358757,0],[0.882142515,0,0,-0.470982573],[0,0,0,0],[9E+09,9E+09,9E+09,9E+09,9E+09,9E+09]];
    CONST robtarget Target_4160:=[[72.726442119,107.1647556,0],[0.882142515,0,0,-0.470982573],[0,0,0,0],[9E+09,9E+09,9E+09,9E+09,9E+09,9E+09]];
    CONST robtarget Target_4170:=[[73.074801243,107.253980112,0],[0.882142515,0,0,-0.470982573],[0,0,0,0],[9E+09,9E+09,9E+09,9E+09,9E+09,9E+09]];
    CONST robtarget Target_4180:=[[73.413608351,107.363032293,0],[0.882142515,0,0,-0.470982573],[0,0,0,0],[9E+09,9E+09,9E+09,9E+09,9E+09,9E+09]];
    CONST robtarget Target_4190:=[[73.742863443,107.491912143,0],[0.882142515,0,0,-0.470982573],[0,0,0,0],[9E+09,9E+09,9E+09,9E+09,9E+09,9E+09]];
    CONST robtarget Target_4200:=[[74.062566519,107.640619663,0],[0.882142515,0,0,-0.470982573],[0,0,0,0],[9E+09,9E+09,9E+09,9E+09,9E+09,9E+09]];
    CONST robtarget Target_4210:=[[74.368809937,107.805970846,0],[0.882142515,0,0,-0.470982573],[0,0,0,0],[9E+09,9E+09,9E+09,9E+09,9E+09,9E+09]];
    CONST robtarget Target_4220:=[[74.657686053,107.984781689,0],[0.882142515,0,0,-0.470982573],[0,0,0,0],[9E+09,9E+09,9E+09,9E+09,9E+09,9E+09]];
    CONST robtarget Target_4230:=[[74.929194867,108.17705219,0],[0.882142515,0,0,-0.470982573],[0,0,0,0],[9E+09,9E+09,9E+09,9E+09,9E+09,9E+09]];
    CONST robtarget Target_4240:=[[75.18333638,108.382782349,0],[0.882142515,0,0,-0.470982573],[0,0,0,0],[9E+09,9E+09,9E+09,9E+09,9E+09,9E+09]];
    CONST robtarget Target_4250:=[[75.420110591,108.601972168,0],[0.882142515,0,0,-0.470982573],[0,0,0,0],[9E+09,9E+09,9E+09,9E+09,9E+09,9E+09]];
    CONST robtarget Target_4260:=[[75.639517501,108.834621645,0],[0.882142515,0,0,-0.470982573],[0,0,0,0],[9E+09,9E+09,9E+09,9E+09,9E+09,9E+09]];
    CONST robtarget Target_4270:=[[75.841557109,109.080730781,0],[0.882142515,0,0,-0.470982573],[0,0,0,0],[9E+09,9E+09,9E+09,9E+09,9E+09,9E+09]];
    CONST robtarget Target_4280:=[[76.026229416,109.340299575,0],[0.882142515,0,0,-0.470982573],[0,0,0,0],[9E+09,9E+09,9E+09,9E+09,9E+09,9E+09]];
    CONST robtarget Target_4290:=[[76.276897468,109.77708721,0],[0.882142515,0,0,-0.470982573],[0,0,0,0],[9E+09,9E+09,9E+09,9E+09,9E+09,9E+09]];
    CONST robtarget Target_4300:=[[76.482410537,110.216769394,0],[0.882142515,0,0,-0.470982573],[0,0,0,0],[9E+09,9E+09,9E+09,9E+09,9E+09,9E+09]];
    CONST robtarget Target_4310:=[[76.642768621,110.659346129,0],[0.882142515,0,0,-0.470982573],[0,0,0,0],[9E+09,9E+09,9E+09,9E+09,9E+09,9E+09]];
    CONST robtarget Target_4320:=[[76.757971721,111.104817414,0],[0.882142515,0,0,-0.470982573],[0,0,0,0],[9E+09,9E+09,9E+09,9E+09,9E+09,9E+09]];
    CONST robtarget Target_4330:=[[76.839019129,111.582707662,0],[0.882142515,0,0,-0.470982573],[0,0,0,0],[9E+09,9E+09,9E+09,9E+09,9E+09,9E+09]];
    CONST robtarget Target_4340:=[[76.896910134,112.122541285,0],[0.882142515,0,0,-0.470982573],[0,0,0,0],[9E+09,9E+09,9E+09,9E+09,9E+09,9E+09]];
    CONST robtarget Target_4350:=[[76.931644737,112.724318284,0],[0.882142515,0,0,-0.470982573],[0,0,0,0],[9E+09,9E+09,9E+09,9E+09,9E+09,9E+09]];
    CONST robtarget Target_4360:=[[76.943222938,113.388038659,0],[0.882142515,0,0,-0.470982573],[0,0,0,0],[9E+09,9E+09,9E+09,9E+09,9E+09,9E+09]];
    CONST robtarget Target_4370:=[[76.943222938,116.018605935,0],[0.882142515,0,0,-0.470982573],[0,0,0,0],[9E+09,9E+09,9E+09,9E+09,9E+09,9E+09]];
    CONST robtarget Target_4380:=[[65.513222871,116.018605935,0],[0.882142515,0,0,-0.470982573],[0,0,0,0],[9E+09,9E+09,9E+09,9E+09,9E+09,9E+09]];
    CONST robtarget Target_4390:=[[75.6279393,114.499545959,0],[0.882142515,0,0,-0.470982573],[0,0,0,0],[9E+09,9E+09,9E+09,9E+09,9E+09,9E+09]];
    CONST robtarget Target_4400:=[[66.828506509,114.499545959,0],[0.882142515,0,0,-0.470982573],[0,0,0,0],[9E+09,9E+09,9E+09,9E+09,9E+09,9E+09]];
    CONST robtarget Target_4410:=[[66.828506509,113.341725855,0],[0.882142515,0,0,-0.470982573],[0,0,0,0],[9E+09,9E+09,9E+09,9E+09,9E+09,9E+09]];
    CONST robtarget Target_4420:=[[66.838637435,112.848783946,0],[0.882142515,0,0,-0.470982573],[0,0,0,0],[9E+09,9E+09,9E+09,9E+09,9E+09,9E+09]];
    CONST robtarget Target_4430:=[[66.869030213,112.39810247,0],[0.882142515,0,0,-0.470982573],[0,0,0,0],[9E+09,9E+09,9E+09,9E+09,9E+09,9E+09]];
    CONST robtarget Target_4440:=[[66.919684843,111.989681428,0],[0.882142515,0,0,-0.470982573],[0,0,0,0],[9E+09,9E+09,9E+09,9E+09,9E+09,9E+09]];
    CONST robtarget Target_4450:=[[66.990601324,111.62352082,0],[0.882142515,0,0,-0.470982573],[0,0,0,0],[9E+09,9E+09,9E+09,9E+09,9E+09,9E+09]];
    CONST robtarget Target_4460:=[[67.084095297,111.283411165,0],[0.882142515,0,0,-0.470982573],[0,0,0,0],[9E+09,9E+09,9E+09,9E+09,9E+09,9E+09]];
    CONST robtarget Target_4470:=[[67.202482403,110.95314298,0],[0.882142515,0,0,-0.470982573],[0,0,0,0],[9E+09,9E+09,9E+09,9E+09,9E+09,9E+09]];
    CONST robtarget Target_4480:=[[67.345762641,110.632716266,0],[0.882142515,0,0,-0.470982573],[0,0,0,0],[9E+09,9E+09,9E+09,9E+09,9E+09,9E+09]];
    CONST robtarget Target_4490:=[[67.513936011,110.322131024,0],[0.882142515,0,0,-0.470982573],[0,0,0,0],[9E+09,9E+09,9E+09,9E+09,9E+09,9E+09]];
    CONST robtarget Target_4500:=[[67.803101582,109.918051807,0],[0.882142515,0,0,-0.470982573],[0,0,0,0],[9E+09,9E+09,9E+09,9E+09,9E+09,9E+09]];
    CONST robtarget Target_4510:=[[68.142632327,109.567232316,0],[0.882142515,0,0,-0.470982573],[0,0,0,0],[9E+09,9E+09,9E+09,9E+09,9E+09,9E+09]];
    CONST robtarget Target_4520:=[[68.532528247,109.269672549,0],[0.882142515,0,0,-0.470982573],[0,0,0,0],[9E+09,9E+09,9E+09,9E+09,9E+09,9E+09]];
    CONST robtarget Target_4530:=[[68.972789342,109.025372507,0],[0.882142515,0,0,-0.470982573],[0,0,0,0],[9E+09,9E+09,9E+09,9E+09,9E+09,9E+09]];
    CONST robtarget Target_4540:=[[69.462257791,108.8349111,0],[0.882142515,0,0,-0.470982573],[0,0,0,0],[9E+09,9E+09,9E+09,9E+09,9E+09,9E+09]];
    CONST robtarget Target_4550:=[[69.999775774,108.698867238,0],[0.882142515,0,0,-0.470982573],[0,0,0,0],[9E+09,9E+09,9E+09,9E+09,9E+09,9E+09]];
    CONST robtarget Target_4560:=[[70.585343292,108.61724092,0],[0.882142515,0,0,-0.470982573],[0,0,0,0],[9E+09,9E+09,9E+09,9E+09,9E+09,9E+09]];
    CONST robtarget Target_4570:=[[71.218960344,108.590032148,0],[0.882142515,0,0,-0.470982573],[0,0,0,0],[9E+09,9E+09,9E+09,9E+09,9E+09,9E+09]];
    CONST robtarget Target_4580:=[[71.858077041,108.61492528,0],[0.882142515,0,0,-0.470982573],[0,0,0,0],[9E+09,9E+09,9E+09,9E+09,9E+09,9E+09]];
    CONST robtarget Target_4590:=[[72.441618374,108.689604677,0],[0.882142515,0,0,-0.470982573],[0,0,0,0],[9E+09,9E+09,9E+09,9E+09,9E+09,9E+09]];
    CONST robtarget Target_4600:=[[72.969584341,108.814070338,0],[0.882142515,0,0,-0.470982573],[0,0,0,0],[9E+09,9E+09,9E+09,9E+09,9E+09,9E+09]];
    CONST robtarget Target_4610:=[[73.441974943,108.988322264,0],[0.882142515,0,0,-0.470982573],[0,0,0,0],[9E+09,9E+09,9E+09,9E+09,9E+09,9E+09]];
    CONST robtarget Target_4620:=[[73.864579281,109.212360454,0],[0.882142515,0,0,-0.470982573],[0,0,0,0],[9E+09,9E+09,9E+09,9E+09,9E+09,9E+09]];
    CONST robtarget Target_4630:=[[74.243186455,109.486184908,0],[0.882142515,0,0,-0.470982573],[0,0,0,0],[9E+09,9E+09,9E+09,9E+09,9E+09,9E+09]];
    CONST robtarget Target_4640:=[[74.577796466,109.809795628,0],[0.882142515,0,0,-0.470982573],[0,0,0,0],[9E+09,9E+09,9E+09,9E+09,9E+09,9E+09]];
    CONST robtarget Target_4650:=[[74.868409312,110.183192611,0],[0.882142515,0,0,-0.470982573],[0,0,0,0],[9E+09,9E+09,9E+09,9E+09,9E+09,9E+09]];
    CONST robtarget Target_4660:=[[75.069001645,110.502461505,0],[0.882142515,0,0,-0.470982573],[0,0,0,0],[9E+09,9E+09,9E+09,9E+09,9E+09,9E+09]];
    CONST robtarget Target_4670:=[[75.235438285,110.83967661,0],[0.882142515,0,0,-0.470982573],[0,0,0,0],[9E+09,9E+09,9E+09,9E+09,9E+09,9E+09]];
    CONST robtarget Target_4680:=[[75.367719231,111.194837927,0],[0.882142515,0,0,-0.470982573],[0,0,0,0],[9E+09,9E+09,9E+09,9E+09,9E+09,9E+09]];
    CONST robtarget Target_4690:=[[75.465844485,111.567945455,0],[0.882142515,0,0,-0.470982573],[0,0,0,0],[9E+09,9E+09,9E+09,9E+09,9E+09,9E+09]];
    CONST robtarget Target_4700:=[[75.536760967,111.965367206,0],[0.882142515,0,0,-0.470982573],[0,0,0,0],[9E+09,9E+09,9E+09,9E+09,9E+09,9E+09]];
    CONST robtarget Target_4710:=[[75.587415596,112.39347119,0],[0.882142515,0,0,-0.470982573],[0,0,0,0],[9E+09,9E+09,9E+09,9E+09,9E+09,9E+09]];
    CONST robtarget Target_4720:=[[75.617808374,112.852257406,0],[0.882142515,0,0,-0.470982573],[0,0,0,0],[9E+09,9E+09,9E+09,9E+09,9E+09,9E+09]];
    CONST robtarget Target_4730:=[[75.6279393,113.341725855,0],[0.882142515,0,0,-0.470982573],[0,0,0,0],[9E+09,9E+09,9E+09,9E+09,9E+09,9E+09]];
    CONST robtarget Target_4740:=[[76.943222938,100.448241177,0],[0.882142515,0,0,-0.470982573],[0,0,0,0],[9E+09,9E+09,9E+09,9E+09,9E+09,9E+09]];
    CONST robtarget Target_4750:=[[76.943222938,98.9291812,0],[0.882142515,0,0,-0.470982573],[0,0,0,0],[9E+09,9E+09,9E+09,9E+09,9E+09,9E+09]];
    CONST robtarget Target_4760:=[[72.395305569,98.9291812,0],[0.882142515,0,0,-0.470982573],[0,0,0,0],[9E+09,9E+09,9E+09,9E+09,9E+09,9E+09]];
    CONST robtarget Target_4770:=[[72.395305569,97.187819764,0],[0.882142515,0,0,-0.470982573],[0,0,0,0],[9E+09,9E+09,9E+09,9E+09,9E+09,9E+09]];
    CONST robtarget Target_4780:=[[76.943222938,93.575421039,0],[0.882142515,0,0,-0.470982573],[0,0,0,0],[9E+09,9E+09,9E+09,9E+09,9E+09,9E+09]];
    CONST robtarget Target_4790:=[[76.943222938,91.602495582,0],[0.882142515,0,0,-0.470982573],[0,0,0,0],[9E+09,9E+09,9E+09,9E+09,9E+09,9E+09]];
    CONST robtarget Target_4800:=[[71.969227771,95.668759787,0],[0.882142515,0,0,-0.470982573],[0,0,0,0],[9E+09,9E+09,9E+09,9E+09,9E+09,9E+09]];
    CONST robtarget Target_4810:=[[71.737953205,95.150635291,0],[0.882142515,0,0,-0.470982573],[0,0,0,0],[9E+09,9E+09,9E+09,9E+09,9E+09,9E+09]];
    CONST robtarget Target_4820:=[[71.451682185,94.689243979,0],[0.882142515,0,0,-0.470982573],[0,0,0,0],[9E+09,9E+09,9E+09,9E+09,9E+09,9E+09]];
    CONST robtarget Target_4830:=[[71.110414709,94.284585853,0],[0.882142515,0,0,-0.470982573],[0,0,0,0],[9E+09,9E+09,9E+09,9E+09,9E+09,9E+09]];
    CONST robtarget Target_4840:=[[70.714150778,93.936660912,0],[0.882142515,0,0,-0.470982573],[0,0,0,0],[9E+09,9E+09,9E+09,9E+09,9E+09,9E+09]];
    CONST robtarget Target_4850:=[[70.495974053,93.786867936,0],[0.882142515,0,0,-0.470982573],[0,0,0,0],[9E+09,9E+09,9E+09,9E+09,9E+09,9E+09]];
    CONST robtarget Target_4860:=[[70.265206033,93.657047357,0],[0.882142515,0,0,-0.470982573],[0,0,0,0],[9E+09,9E+09,9E+09,9E+09,9E+09,9E+09]];
    CONST robtarget Target_4870:=[[70.02184672,93.547199174,0],[0.882142515,0,0,-0.470982573],[0,0,0,0],[9E+09,9E+09,9E+09,9E+09,9E+09,9E+09]];
    CONST robtarget Target_4880:=[[69.765896113,93.457323389,0],[0.882142515,0,0,-0.470982573],[0,0,0,0],[9E+09,9E+09,9E+09,9E+09,9E+09,9E+09]];
    CONST robtarget Target_4890:=[[69.497354213,93.38742,0],[0.882142515,0,0,-0.470982573],[0,0,0,0],[9E+09,9E+09,9E+09,9E+09,9E+09,9E+09]];
    CONST robtarget Target_4900:=[[69.216221019,93.337489008,0],[0.882142515,0,0,-0.470982573],[0,0,0,0],[9E+09,9E+09,9E+09,9E+09,9E+09,9E+09]];
    CONST robtarget Target_4910:=[[68.922496531,93.307530413,0],[0.882142515,0,0,-0.470982573],[0,0,0,0],[9E+09,9E+09,9E+09,9E+09,9E+09,9E+09]];
    CONST robtarget Target_4920:=[[68.61618075,93.297544214,0],[0.882142515,0,0,-0.470982573],[0,0,0,0],[9E+09,9E+09,9E+09,9E+09,9E+09,9E+09]];
    CONST robtarget Target_4930:=[[68.185182216,93.319253341,0],[0.882142515,0,0,-0.470982573],[0,0,0,0],[9E+09,9E+09,9E+09,9E+09,9E+09,9E+09]];
    CONST robtarget Target_4940:=[[67.790655016,93.384380722,0],[0.882142515,0,0,-0.470982573],[0,0,0,0],[9E+09,9E+09,9E+09,9E+09,9E+09,9E+09]];
    CONST robtarget Target_4950:=[[67.432599149,93.492926357,0],[0.882142515,0,0,-0.470982573],[0,0,0,0],[9E+09,9E+09,9E+09,9E+09,9E+09,9E+09]];
    CONST robtarget Target_4960:=[[67.111014615,93.644890245,0],[0.882142515,0,0,-0.470982573],[0,0,0,0],[9E+09,9E+09,9E+09,9E+09,9E+09,9E+09]];
    CONST robtarget Target_4970:=[[66.821270134,93.834483287,0],[0.882142515,0,0,-0.470982573],[0,0,0,0],[9E+09,9E+09,9E+09,9E+09,9E+09,9E+09]];
    CONST robtarget Target_4980:=[[66.558734425,94.055916382,0],[0.882142515,0,0,-0.470982573],[0,0,0,0],[9E+09,9E+09,9E+09,9E+09,9E+09,9E+09]];
    CONST robtarget Target_4990:=[[66.323407489,94.30918953,0],[0.882142515,0,0,-0.470982573],[0,0,0,0],[9E+09,9E+09,9E+09,9E+09,9E+09,9E+09]];
    CONST robtarget Target_5000:=[[66.115289325,94.594302731,0],[0.882142515,0,0,-0.470982573],[0,0,0,0],[9E+09,9E+09,9E+09,9E+09,9E+09,9E+09]];
    CONST robtarget Target_5010:=[[65.938432304,94.899098873,0],[0.882142515,0,0,-0.470982573],[0,0,0,0],[9E+09,9E+09,9E+09,9E+09,9E+09,9E+09]];
    CONST robtarget Target_5020:=[[65.796888797,95.211420846,0],[0.882142515,0,0,-0.470982573],[0,0,0,0],[9E+09,9E+09,9E+09,9E+09,9E+09,9E+09]];
    CONST robtarget Target_5030:=[[65.690658802,95.53126865,0],[0.882142515,0,0,-0.470982573],[0,0,0,0],[9E+09,9E+09,9E+09,9E+09,9E+09,9E+09]];
    CONST robtarget Target_5040:=[[65.619742321,95.858642284,0],[0.882142515,0,0,-0.470982573],[0,0,0,0],[9E+09,9E+09,9E+09,9E+09,9E+09,9E+09]];
    CONST robtarget Target_5050:=[[65.573140062,96.209751231,0],[0.882142515,0,0,-0.470982573],[0,0,0,0],[9E+09,9E+09,9E+09,9E+09,9E+09,9E+09]];
    CONST robtarget Target_5060:=[[65.539852734,96.600804971,0],[0.882142515,0,0,-0.470982573],[0,0,0,0],[9E+09,9E+09,9E+09,9E+09,9E+09,9E+09]];
    CONST robtarget Target_5070:=[[65.519880337,97.031803505,0],[0.882142515,0,0,-0.470982573],[0,0,0,0],[9E+09,9E+09,9E+09,9E+09,9E+09,9E+09]];
    CONST robtarget Target_5080:=[[65.513222871,97.502746832,0],[0.882142515,0,0,-0.470982573],[0,0,0,0],[9E+09,9E+09,9E+09,9E+09,9E+09,9E+09]];
    CONST robtarget Target_5090:=[[65.513222871,100.448241177,0],[0.882142515,0,0,-0.470982573],[0,0,0,0],[9E+09,9E+09,9E+09,9E+09,9E+09,9E+09]];
    CONST robtarget Target_5100:=[[76.943222938,100.448241177,0],[0.882142515,0,0,-0.470982573],[0,0,0,0],[9E+09,9E+09,9E+09,9E+09,9E+09,9E+09]];
    CONST robtarget Target_5110:=[[71.126334735,98.9291812,0],[0.882142515,0,0,-0.470982573],[0,0,0,0],[9E+09,9E+09,9E+09,9E+09,9E+09,9E+09]];
    CONST robtarget Target_5120:=[[71.126334735,97.59537244,0],[0.882142515,0,0,-0.470982573],[0,0,0,0],[9E+09,9E+09,9E+09,9E+09,9E+09,9E+09]];
    CONST robtarget Target_5130:=[[71.11909836,97.274945727,0],[0.882142515,0,0,-0.470982573],[0,0,0,0],[9E+09,9E+09,9E+09,9E+09,9E+09,9E+09]];
    CONST robtarget Target_5140:=[[71.097389233,96.971307404,0],[0.882142515,0,0,-0.470982573],[0,0,0,0],[9E+09,9E+09,9E+09,9E+09,9E+09,9E+09]];
    CONST robtarget Target_5150:=[[71.061207355,96.684457473,0],[0.882142515,0,0,-0.470982573],[0,0,0,0],[9E+09,9E+09,9E+09,9E+09,9E+09,9E+09]];
    CONST robtarget Target_5160:=[[71.010552725,96.414395934,0],[0.882142515,0,0,-0.470982573],[0,0,0,0],[9E+09,9E+09,9E+09,9E+09,9E+09,9E+09]];
    CONST robtarget Target_5170:=[[70.937320604,96.162859517,0],[0.882142515,0,0,-0.470982573],[0,0,0,0],[9E+09,9E+09,9E+09,9E+09,9E+09,9E+09]];
    CONST robtarget Target_5180:=[[70.833406249,95.931584951,0],[0.882142515,0,0,-0.470982573],[0,0,0,0],[9E+09,9E+09,9E+09,9E+09,9E+09,9E+09]];
    CONST robtarget Target_5190:=[[70.698809662,95.720572237,0],[0.882142515,0,0,-0.470982573],[0,0,0,0],[9E+09,9E+09,9E+09,9E+09,9E+09,9E+09]];
    CONST robtarget Target_5200:=[[70.533530842,95.529821375,0],[0.882142515,0,0,-0.470982573],[0,0,0,0],[9E+09,9E+09,9E+09,9E+09,9E+09,9E+09]];
    CONST robtarget Target_5210:=[[70.367962567,95.374094571,0],[0.882142515,0,0,-0.470982573],[0,0,0,0],[9E+09,9E+09,9E+09,9E+09,9E+09,9E+09]];
    CONST robtarget Target_5220:=[[70.186184811,95.240366349,0],[0.882142515,0,0,-0.470982573],[0,0,0,0],[9E+09,9E+09,9E+09,9E+09,9E+09,9E+09]];
    CONST robtarget Target_5230:=[[69.988197573,95.128636709,0],[0.882142515,0,0,-0.470982573],[0,0,0,0],[9E+09,9E+09,9E+09,9E+09,9E+09,9E+09]];
    CONST robtarget Target_5240:=[[69.774000854,95.038905651,0],[0.882142515,0,0,-0.470982573],[0,0,0,0],[9E+09,9E+09,9E+09,9E+09,9E+09,9E+09]];
    CONST robtarget Target_5250:=[[69.542436833,94.970015354,0],[0.882142515,0,0,-0.470982573],[0,0,0,0],[9E+09,9E+09,9E+09,9E+09,9E+09,9E+09]];
    CONST robtarget Target_5260:=[[69.292347691,94.920808,0],[0.882142515,0,0,-0.470982573],[0,0,0,0],[9E+09,9E+09,9E+09,9E+09,9E+09,9E+09]];
    CONST robtarget Target_5270:=[[69.023733427,94.891283587,0],[0.882142515,0,0,-0.470982573],[0,0,0,0],[9E+09,9E+09,9E+09,9E+09,9E+09,9E+09]];
    CONST robtarget Target_5280:=[[68.736594041,94.881442117,0],[0.882142515,0,0,-0.470982573],[0,0,0,0],[9E+09,9E+09,9E+09,9E+09,9E+09,9E+09]];
    CONST robtarget Target_5290:=[[68.493741274,94.892441408,0],[0.882142515,0,0,-0.470982573],[0,0,0,0],[9E+09,9E+09,9E+09,9E+09,9E+09,9E+09]];
    CONST robtarget Target_5300:=[[68.265361258,94.92543928,0],[0.882142515,0,0,-0.470982573],[0,0,0,0],[9E+09,9E+09,9E+09,9E+09,9E+09,9E+09]];
    CONST robtarget Target_5310:=[[68.051453994,94.980435735,0],[0.882142515,0,0,-0.470982573],[0,0,0,0],[9E+09,9E+09,9E+09,9E+09,9E+09,9E+09]];
    CONST robtarget Target_5320:=[[67.852019481,95.057430772,0],[0.882142515,0,0,-0.470982573],[0,0,0,0],[9E+09,9E+09,9E+09,9E+09,9E+09,9E+09]];
    CONST robtarget Target_5330:=[[67.66821554,95.157582211,0],[0.882142515,0,0,-0.470982573],[0,0,0,0],[9E+09,9E+09,9E+09,9E+09,9E+09,9E+09]];
    CONST robtarget Target_5340:=[[67.50119999,95.282047873,0],[0.882142515,0,0,-0.470982573],[0,0,0,0],[9E+09,9E+09,9E+09,9E+09,9E+09,9E+09]];
    CONST robtarget Target_5350:=[[67.350972831,95.430827756,0],[0.882142515,0,0,-0.470982573],[0,0,0,0],[9E+09,9E+09,9E+09,9E+09,9E+09,9E+09]];
    CONST robtarget Target_5360:=[[67.217534064,95.603921861,0],[0.882142515,0,0,-0.470982573],[0,0,0,0],[9E+09,9E+09,9E+09,9E+09,9E+09,9E+09]];
    CONST robtarget Target_5370:=[[67.1188299,95.772674142,0],[0.882142515,0,0,-0.470982573],[0,0,0,0],[9E+09,9E+09,9E+09,9E+09,9E+09,9E+09]];
    CONST robtarget Target_5380:=[[67.035756308,95.954741353,0],[0.882142515,0,0,-0.470982573],[0,0,0,0],[9E+09,9E+09,9E+09,9E+09,9E+09,9E+09]];
    CONST robtarget Target_5390:=[[66.968313287,96.150123495,0],[0.882142515,0,0,-0.470982573],[0,0,0,0],[9E+09,9E+09,9E+09,9E+09,9E+09,9E+09]];
    CONST robtarget Target_5400:=[[66.916500837,96.358820569,0],[0.882142515,0,0,-0.470982573],[0,0,0,0],[9E+09,9E+09,9E+09,9E+09,9E+09,9E+09]];
    CONST robtarget Target_5410:=[[66.878003319,96.586621675,0],[0.882142515,0,0,-0.470982573],[0,0,0,0],[9E+09,9E+09,9E+09,9E+09,9E+09,9E+09]];
    CONST robtarget Target_5420:=[[66.850505091,96.839315912,0],[0.882142515,0,0,-0.470982573],[0,0,0,0],[9E+09,9E+09,9E+09,9E+09,9E+09,9E+09]];
    CONST robtarget Target_5430:=[[66.834006155,97.116903282,0],[0.882142515,0,0,-0.470982573],[0,0,0,0],[9E+09,9E+09,9E+09,9E+09,9E+09,9E+09]];
    CONST robtarget Target_5440:=[[66.828506509,97.419383785,0],[0.882142515,0,0,-0.470982573],[0,0,0,0],[9E+09,9E+09,9E+09,9E+09,9E+09,9E+09]];
    CONST robtarget Target_5450:=[[66.828506509,98.9291812,0],[0.882142515,0,0,-0.470982573],[0,0,0,0],[9E+09,9E+09,9E+09,9E+09,9E+09,9E+09]];
    CONST robtarget Target_5460:=[[71.126334735,98.9291812,0],[0.882142515,0,0,-0.470982573],[0,0,0,0],[9E+09,9E+09,9E+09,9E+09,9E+09,9E+09]];
    CONST robtarget Target_5470:=[[70.832489087,106.240000104,-227.23325525],[0.882142515,0,0,-0.470982573],[0,-1,0,0],[9E+09,9E+09,9E+09,9E+09,9E+09,9E+09]];
    CONST robtarget Target_5480:=[[65.513222871,89.314643056,0],[0.882142515,0,0,-0.470982573],[0,0,0,0],[9E+09,9E+09,9E+09,9E+09,9E+09,9E+09]];
    CONST robtarget Target_5490:=[[65.513222871,90.833703033,0],[0.882142515,0,0,-0.470982573],[0,0,0,0],[9E+09,9E+09,9E+09,9E+09,9E+09,9E+09]];
    CONST robtarget Target_5500:=[[72.645394712,90.833703033,0],[0.882142515,0,0,-0.470982573],[0,0,0,0],[9E+09,9E+09,9E+09,9E+09,9E+09,9E+09]];
    CONST robtarget Target_5510:=[[73.232409505,90.818361917,0],[0.882142515,0,0,-0.470982573],[0,0,0,0],[9E+09,9E+09,9E+09,9E+09,9E+09,9E+09]];
    CONST robtarget Target_5520:=[[73.770795853,90.772338567,0],[0.882142515,0,0,-0.470982573],[0,0,0,0],[9E+09,9E+09,9E+09,9E+09,9E+09,9E+09]];
    CONST robtarget Target_5530:=[[74.260553757,90.695632986,0],[0.882142515,0,0,-0.470982573],[0,0,0,0],[9E+09,9E+09,9E+09,9E+09,9E+09,9E+09]];
    CONST robtarget Target_5540:=[[74.701683217,90.588245171,0],[0.882142515,0,0,-0.470982573],[0,0,0,0],[9E+09,9E+09,9E+09,9E+09,9E+09,9E+09]];
    CONST robtarget Target_5550:=[[75.103446793,90.443228203,0],[0.882142515,0,0,-0.470982573],[0,0,0,0],[9E+09,9E+09,9E+09,9E+09,9E+09,9E+09]];
    CONST robtarget Target_5560:=[[75.475107046,90.253635161,0],[0.882142515,0,0,-0.470982573],[0,0,0,0],[9E+09,9E+09,9E+09,9E+09,9E+09,9E+09]];
    CONST robtarget Target_5570:=[[75.816663977,90.019466045,0],[0.882142515,0,0,-0.470982573],[0,0,0,0],[9E+09,9E+09,9E+09,9E+09,9E+09,9E+09]];
    CONST robtarget Target_5580:=[[76.128117585,89.740720855,0],[0.882142515,0,0,-0.470982573],[0,0,0,0],[9E+09,9E+09,9E+09,9E+09,9E+09,9E+09]];
    CONST robtarget Target_5590:=[[76.375601632,89.46284403,0],[0.882142515,0,0,-0.470982573],[0,0,0,0],[9E+09,9E+09,9E+09,9E+09,9E+09,9E+09]];
    CONST robtarget Target_5600:=[[76.590087806,89.157179522,0],[0.882142515,0,0,-0.470982573],[0,0,0,0],[9E+09,9E+09,9E+09,9E+09,9E+09,9E+09]];
    CONST robtarget Target_5610:=[[76.771576108,88.823727332,0],[0.882142515,0,0,-0.470982573],[0,0,0,0],[9E+09,9E+09,9E+09,9E+09,9E+09,9E+09]];
    CONST robtarget Target_5620:=[[76.920066536,88.46248746,0],[0.882142515,0,0,-0.470982573],[0,0,0,0],[9E+09,9E+09,9E+09,9E+09,9E+09,9E+09]];
    CONST robtarget Target_5630:=[[77.035559091,88.071144265,0],[0.882142515,0,0,-0.470982573],[0,0,0,0],[9E+09,9E+09,9E+09,9E+09,9E+09,9E+09]];
    CONST robtarget Target_5640:=[[77.118053774,87.647382107,0],[0.882142515,0,0,-0.470982573],[0,0,0,0],[9E+09,9E+09,9E+09,9E+09,9E+09,9E+09]];
    CONST robtarget Target_5650:=[[77.167550583,87.191200986,0],[0.882142515,0,0,-0.470982573],[0,0,0,0],[9E+09,9E+09,9E+09,9E+09,9E+09,9E+09]];
    CONST robtarget Target_5660:=[[77.18404952,86.702600902,0],[0.882142515,0,0,-0.470982573],[0,0,0,0],[9E+09,9E+09,9E+09,9E+09,9E+09,9E+09]];
    CONST robtarget Target_5670:=[[77.167840038,86.195475696,0],[0.882142515,0,0,-0.470982573],[0,0,0,0],[9E+09,9E+09,9E+09,9E+09,9E+09,9E+09]];
    CONST robtarget Target_5680:=[[77.119211594,85.730032014,0],[0.882142515,0,0,-0.470982573],[0,0,0,0],[9E+09,9E+09,9E+09,9E+09,9E+09,9E+09]];
    CONST robtarget Target_5690:=[[77.038164187,85.306269856,0],[0.882142515,0,0,-0.470982573],[0,0,0,0],[9E+09,9E+09,9E+09,9E+09,9E+09,9E+09]];
    CONST robtarget Target_5700:=[[76.924697816,84.924189222,0],[0.882142515,0,0,-0.470982573],[0,0,0,0],[9E+09,9E+09,9E+09,9E+09,9E+09,9E+09]];
    CONST robtarget Target_5710:=[[76.777654663,84.573948641,0],[0.882142515,0,0,-0.470982573],[0,0,0,0],[9E+09,9E+09,9E+09,9E+09,9E+09,9E+09]];
    CONST robtarget Target_5720:=[[76.595876907,84.245706641,0],[0.882142515,0,0,-0.470982573],[0,0,0,0],[9E+09,9E+09,9E+09,9E+09,9E+09,9E+09]];
    CONST robtarget Target_5730:=[[76.379364547,83.939463224,0],[0.882142515,0,0,-0.470982573],[0,0,0,0],[9E+09,9E+09,9E+09,9E+09,9E+09,9E+09]];
    CONST robtarget Target_5740:=[[76.128117585,83.655218388,0],[0.882142515,0,0,-0.470982573],[0,0,0,0],[9E+09,9E+09,9E+09,9E+09,9E+09,9E+09]];
    CONST robtarget Target_5750:=[[75.819558527,83.372710283,0],[0.882142515,0,0,-0.470982573],[0,0,0,0],[9E+09,9E+09,9E+09,9E+09,9E+09,9E+09]];
    CONST robtarget Target_5760:=[[75.477422686,83.136514981,0],[0.882142515,0,0,-0.470982573],[0,0,0,0],[9E+09,9E+09,9E+09,9E+09,9E+09,9E+09]];
    CONST robtarget Target_5770:=[[75.101710063,82.946632484,0],[0.882142515,0,0,-0.470982573],[0,0,0,0],[9E+09,9E+09,9E+09,9E+09,9E+09,9E+09]];
    CONST robtarget Target_5780:=[[74.692420656,82.803062792,0],[0.882142515,0,0,-0.470982573],[0,0,0,0],[9E+09,9E+09,9E+09,9E+09,9E+09,9E+09]];
    CONST robtarget Target_5790:=[[74.244923186,82.697701162,0],[0.882142515,0,0,-0.470982573],[0,0,0,0],[9E+09,9E+09,9E+09,9E+09,9E+09,9E+09]];
    CONST robtarget Target_5800:=[[73.754586372,82.622442855,0],[0.882142515,0,0,-0.470982573],[0,0,0,0],[9E+09,9E+09,9E+09,9E+09,9E+09,9E+09]];
    CONST robtarget Target_5810:=[[73.221410214,82.577287871,0],[0.882142515,0,0,-0.470982573],[0,0,0,0],[9E+09,9E+09,9E+09,9E+09,9E+09,9E+09]];
    CONST robtarget Target_5820:=[[72.645394712,82.56223621,0],[0.882142515,0,0,-0.470982573],[0,0,0,0],[9E+09,9E+09,9E+09,9E+09,9E+09,9E+09]];
    CONST robtarget Target_5830:=[[65.513222871,82.56223621,0],[0.882142515,0,0,-0.470982573],[0,0,0,0],[9E+09,9E+09,9E+09,9E+09,9E+09,9E+09]];
    CONST robtarget Target_5840:=[[65.513222871,84.081296186,0],[0.882142515,0,0,-0.470982573],[0,0,0,0],[9E+09,9E+09,9E+09,9E+09,9E+09,9E+09]];
    CONST robtarget Target_5850:=[[72.682444955,84.081296186,0],[0.882142515,0,0,-0.470982573],[0,0,0,0],[9E+09,9E+09,9E+09,9E+09,9E+09,9E+09]];
    CONST robtarget Target_5860:=[[73.052079023,84.087664197,0],[0.882142515,0,0,-0.470982573],[0,0,0,0],[9E+09,9E+09,9E+09,9E+09,9E+09,9E+09]];
    CONST robtarget Target_5870:=[[73.392188679,84.106768229,0],[0.882142515,0,0,-0.470982573],[0,0,0,0],[9E+09,9E+09,9E+09,9E+09,9E+09,9E+09]];
    CONST robtarget Target_5880:=[[73.702773922,84.138608281,0],[0.882142515,0,0,-0.470982573],[0,0,0,0],[9E+09,9E+09,9E+09,9E+09,9E+09,9E+09]];
    CONST robtarget Target_5890:=[[73.983834752,84.183184356,0],[0.882142515,0,0,-0.470982573],[0,0,0,0],[9E+09,9E+09,9E+09,9E+09,9E+09,9E+09]];
    CONST robtarget Target_5900:=[[74.244054821,84.245706641,0],[0.882142515,0,0,-0.470982573],[0,0,0,0],[9E+09,9E+09,9E+09,9E+09,9E+09,9E+09]];
    CONST robtarget Target_5910:=[[74.492117778,84.331385329,0],[0.882142515,0,0,-0.470982573],[0,0,0,0],[9E+09,9E+09,9E+09,9E+09,9E+09,9E+09]];
    CONST robtarget Target_5920:=[[74.728023624,84.440220419,0],[0.882142515,0,0,-0.470982573],[0,0,0,0],[9E+09,9E+09,9E+09,9E+09,9E+09,9E+09]];
    CONST robtarget Target_5930:=[[74.951772359,84.57221191,0],[0.882142515,0,0,-0.470982573],[0,0,0,0],[9E+09,9E+09,9E+09,9E+09,9E+09,9E+09]];
    CONST robtarget Target_5940:=[[75.169153084,84.740674736,0],[0.882142515,0,0,-0.470982573],[0,0,0,0],[9E+09,9E+09,9E+09,9E+09,9E+09,9E+09]];
    CONST robtarget Target_5950:=[[75.358167216,84.940398704,0],[0.882142515,0,0,-0.470982573],[0,0,0,0],[9E+09,9E+09,9E+09,9E+09,9E+09,9E+09]];
    CONST robtarget Target_5960:=[[75.518814755,85.171383814,0],[0.882142515,0,0,-0.470982573],[0,0,0,0],[9E+09,9E+09,9E+09,9E+09,9E+09,9E+09]];
    CONST robtarget Target_5970:=[[75.651095702,85.433630068,0],[0.882142515,0,0,-0.470982573],[0,0,0,0],[9E+09,9E+09,9E+09,9E+09,9E+09,9E+09]];
    CONST robtarget Target_5980:=[[75.754431146,85.721348364,0],[0.882142515,0,0,-0.470982573],[0,0,0,0],[9E+09,9E+09,9E+09,9E+09,9E+09,9E+09]];
    CONST robtarget Target_5990:=[[75.828242178,86.028749601,0],[0.882142515,0,0,-0.470982573],[0,0,0,0],[9E+09,9E+09,9E+09,9E+09,9E+09,9E+09]];
    CONST robtarget Target_6000:=[[75.872528797,86.355833781,0],[0.882142515,0,0,-0.470982573],[0,0,0,0],[9E+09,9E+09,9E+09,9E+09,9E+09,9E+09]];
    CONST robtarget Target_6010:=[[75.887291003,86.702600902,0],[0.882142515,0,0,-0.470982573],[0,0,0,0],[9E+09,9E+09,9E+09,9E+09,9E+09,9E+09]];
    CONST robtarget Target_6020:=[[75.872528797,87.067893145,0],[0.882142515,0,0,-0.470982573],[0,0,0,0],[9E+09,9E+09,9E+09,9E+09,9E+09,9E+09]];
    CONST robtarget Target_6030:=[[75.828242178,87.404239885,0],[0.882142515,0,0,-0.470982573],[0,0,0,0],[9E+09,9E+09,9E+09,9E+09,9E+09,9E+09]];
    CONST robtarget Target_6040:=[[75.754431146,87.711641122,0],[0.882142515,0,0,-0.470982573],[0,0,0,0],[9E+09,9E+09,9E+09,9E+09,9E+09,9E+09]];
    CONST robtarget Target_6050:=[[75.651095702,87.990096857,0],[0.882142515,0,0,-0.470982573],[0,0,0,0],[9E+09,9E+09,9E+09,9E+09,9E+09,9E+09]];
    CONST robtarget Target_6060:=[[75.518814755,88.240186,0],[0.882142515,0,0,-0.470982573],[0,0,0,0],[9E+09,9E+09,9E+09,9E+09,9E+09,9E+09]];
    CONST robtarget Target_6070:=[[75.358167216,88.46248746,0],[0.882142515,0,0,-0.470982573],[0,0,0,0],[9E+09,9E+09,9E+09,9E+09,9E+09,9E+09]];
    CONST robtarget Target_6080:=[[75.169153084,88.657001237,0],[0.882142515,0,0,-0.470982573],[0,0,0,0],[9E+09,9E+09,9E+09,9E+09,9E+09,9E+09]];
    CONST robtarget Target_6090:=[[74.951772359,88.823727332,0],[0.882142515,0,0,-0.470982573],[0,0,0,0],[9E+09,9E+09,9E+09,9E+09,9E+09,9E+09]];
    CONST robtarget Target_6100:=[[74.727734169,88.955718824,0],[0.882142515,0,0,-0.470982573],[0,0,0,0],[9E+09,9E+09,9E+09,9E+09,9E+09,9E+09]];
    CONST robtarget Target_6110:=[[74.490959958,89.064553914,0],[0.882142515,0,0,-0.470982573],[0,0,0,0],[9E+09,9E+09,9E+09,9E+09,9E+09,9E+09]];
    CONST robtarget Target_6120:=[[74.241449725,89.150232602,0],[0.882142515,0,0,-0.470982573],[0,0,0,0],[9E+09,9E+09,9E+09,9E+09,9E+09,9E+09]];
    CONST robtarget Target_6130:=[[73.979203472,89.212754887,0],[0.882142515,0,0,-0.470982573],[0,0,0,0],[9E+09,9E+09,9E+09,9E+09,9E+09,9E+09]];
    CONST robtarget Target_6140:=[[73.694379726,89.257330961,0],[0.882142515,0,0,-0.470982573],[0,0,0,0],[9E+09,9E+09,9E+09,9E+09,9E+09,9E+09]];
    CONST robtarget Target_6150:=[[73.377137018,89.289171014,0],[0.882142515,0,0,-0.470982573],[0,0,0,0],[9E+09,9E+09,9E+09,9E+09,9E+09,9E+09]];
    CONST robtarget Target_6160:=[[73.027475346,89.308275046,0],[0.882142515,0,0,-0.470982573],[0,0,0,0],[9E+09,9E+09,9E+09,9E+09,9E+09,9E+09]];
    CONST robtarget Target_6170:=[[72.645394712,89.314643056,0],[0.882142515,0,0,-0.470982573],[0,0,0,0],[9E+09,9E+09,9E+09,9E+09,9E+09,9E+09]];
    CONST robtarget Target_6180:=[[65.513222871,89.314643056,0],[0.882142515,0,0,-0.470982573],[0,0,0,0],[9E+09,9E+09,9E+09,9E+09,9E+09,9E+09]];
    CONST robtarget Target_6190:=[[65.513222871,76.402633257,0],[0.882142515,0,0,-0.470982573],[0,0,0,0],[9E+09,9E+09,9E+09,9E+09,9E+09,9E+09]];
    CONST robtarget Target_6200:=[[65.513222871,80.830137334,0],[0.882142515,0,0,-0.470982573],[0,0,0,0],[9E+09,9E+09,9E+09,9E+09,9E+09,9E+09]];
    CONST robtarget Target_6210:=[[66.680305536,80.830137334,0],[0.882142515,0,0,-0.470982573],[0,0,0,0],[9E+09,9E+09,9E+09,9E+09,9E+09,9E+09]];
    CONST robtarget Target_6220:=[[66.680305536,79.375915284,0],[0.882142515,0,0,-0.470982573],[0,0,0,0],[9E+09,9E+09,9E+09,9E+09,9E+09,9E+09]];
    CONST robtarget Target_6230:=[[75.776140273,79.375915284,0],[0.882142515,0,0,-0.470982573],[0,0,0,0],[9E+09,9E+09,9E+09,9E+09,9E+09,9E+09]];
    CONST robtarget Target_6240:=[[75.776140273,80.830137334,0],[0.882142515,0,0,-0.470982573],[0,0,0,0],[9E+09,9E+09,9E+09,9E+09,9E+09,9E+09]];
    CONST robtarget Target_6250:=[[76.943222938,80.830137334,0],[0.882142515,0,0,-0.470982573],[0,0,0,0],[9E+09,9E+09,9E+09,9E+09,9E+09,9E+09]];
    CONST robtarget Target_6260:=[[76.943222938,76.402633257,0],[0.882142515,0,0,-0.470982573],[0,0,0,0],[9E+09,9E+09,9E+09,9E+09,9E+09,9E+09]];
    CONST robtarget Target_6270:=[[75.776140273,76.402633257,0],[0.882142515,0,0,-0.470982573],[0,0,0,0],[9E+09,9E+09,9E+09,9E+09,9E+09,9E+09]];
    CONST robtarget Target_6280:=[[75.776140273,77.856855307,0],[0.882142515,0,0,-0.470982573],[0,0,0,0],[9E+09,9E+09,9E+09,9E+09,9E+09,9E+09]];
    CONST robtarget Target_6290:=[[66.680305536,77.856855307,0],[0.882142515,0,0,-0.470982573],[0,0,0,0],[9E+09,9E+09,9E+09,9E+09,9E+09,9E+09]];
    CONST robtarget Target_6300:=[[66.680305536,76.402633257,0],[0.882142515,0,0,-0.470982573],[0,0,0,0],[9E+09,9E+09,9E+09,9E+09,9E+09,9E+09]];
    CONST robtarget Target_6310:=[[65.513222871,76.402633257,0],[0.882142515,0,0,-0.470982573],[0,0,0,0],[9E+09,9E+09,9E+09,9E+09,9E+09,9E+09]];
    CONST robtarget Target_6320:=[[66.865556753,74.939148645,0],[0.882142515,0,0,-0.470982573],[0,0,0,0],[9E+09,9E+09,9E+09,9E+09,9E+09,9E+09]];
    CONST robtarget Target_6330:=[[65.513222871,74.939148645,0],[0.882142515,0,0,-0.470982573],[0,0,0,0],[9E+09,9E+09,9E+09,9E+09,9E+09,9E+09]];
    CONST robtarget Target_6340:=[[65.513222871,67.390161567,0],[0.882142515,0,0,-0.470982573],[0,0,0,0],[9E+09,9E+09,9E+09,9E+09,9E+09,9E+09]];
    CONST robtarget Target_6350:=[[66.884081874,67.390161567,0],[0.882142515,0,0,-0.470982573],[0,0,0,0],[9E+09,9E+09,9E+09,9E+09,9E+09,9E+09]];
    CONST robtarget Target_6360:=[[75.590889057,73.568289642,0],[0.882142515,0,0,-0.470982573],[0,0,0,0],[9E+09,9E+09,9E+09,9E+09,9E+09,9E+09]];
    CONST robtarget Target_6370:=[[75.590889057,67.232698033,0],[0.882142515,0,0,-0.470982573],[0,0,0,0],[9E+09,9E+09,9E+09,9E+09,9E+09,9E+09]];
    CONST robtarget Target_6380:=[[76.943222938,67.232698033,0],[0.882142515,0,0,-0.470982573],[0,0,0,0],[9E+09,9E+09,9E+09,9E+09,9E+09,9E+09]];
    CONST robtarget Target_6390:=[[76.943222938,75.21702547,0],[0.882142515,0,0,-0.470982573],[0,0,0,0],[9E+09,9E+09,9E+09,9E+09,9E+09,9E+09]];
    CONST robtarget Target_6400:=[[75.526051131,75.21702547,0],[0.882142515,0,0,-0.470982573],[0,0,0,0],[9E+09,9E+09,9E+09,9E+09,9E+09,9E+09]];
    CONST robtarget Target_6410:=[[66.865556753,69.103735321,0],[0.882142515,0,0,-0.470982573],[0,0,0,0],[9E+09,9E+09,9E+09,9E+09,9E+09,9E+09]];
    CONST robtarget Target_6420:=[[66.865556753,74.939148645,0],[0.882142515,0,0,-0.470982573],[0,0,0,0],[9E+09,9E+09,9E+09,9E+09,9E+09,9E+09]];
    CONST robtarget Target_6430:=[[95.762416778,129.704038882,0],[0.882142515,0,0,-0.470982573],[0,0,0,0],[9E+09,9E+09,9E+09,9E+09,9E+09,9E+09]];
    CONST robtarget Target_6440:=[[84.332416711,125.850813576,0],[0.882142515,0,0,-0.470982573],[0,0,0,0],[9E+09,9E+09,9E+09,9E+09,9E+09,9E+09]];
    CONST robtarget Target_6450:=[[84.332416711,123.979776288,0],[0.882142515,0,0,-0.470982573],[0,0,0,0],[9E+09,9E+09,9E+09,9E+09,9E+09,9E+09]];
    CONST robtarget Target_6460:=[[95.762416778,120.126550982,0],[0.882142515,0,0,-0.470982573],[0,0,0,0],[9E+09,9E+09,9E+09,9E+09,9E+09,9E+09]];
    CONST robtarget Target_6470:=[[95.762416778,121.728974006,0],[0.882142515,0,0,-0.470982573],[0,0,0,0],[9E+09,9E+09,9E+09,9E+09,9E+09,9E+09]];
    CONST robtarget Target_6480:=[[92.566833291,122.766380819,0],[0.882142515,0,0,-0.470982573],[0,0,0,0],[9E+09,9E+09,9E+09,9E+09,9E+09,9E+09]];
    CONST robtarget Target_6490:=[[92.566833291,127.129046971,0],[0.882142515,0,0,-0.470982573],[0,0,0,0],[9E+09,9E+09,9E+09,9E+09,9E+09,9E+09]];
    CONST robtarget Target_6500:=[[95.762416778,128.166453784,0],[0.882142515,0,0,-0.470982573],[0,0,0,0],[9E+09,9E+09,9E+09,9E+09,9E+09,9E+09]];
    CONST robtarget Target_6510:=[[95.762416778,129.704038882,0],[0.882142515,0,0,-0.470982573],[0,0,0,0],[9E+09,9E+09,9E+09,9E+09,9E+09,9E+09]];
    CONST robtarget Target_6520:=[[91.270074774,126.712231733,0],[0.882142515,0,0,-0.470982573],[0,0,0,0],[9E+09,9E+09,9E+09,9E+09,9E+09,9E+09]];
    CONST robtarget Target_6530:=[[85.888526931,124.952345175,0],[0.882142515,0,0,-0.470982573],[0,0,0,0],[9E+09,9E+09,9E+09,9E+09,9E+09,9E+09]];
    CONST robtarget Target_6540:=[[91.270074774,123.183196056,0],[0.882142515,0,0,-0.470982573],[0,0,0,0],[9E+09,9E+09,9E+09,9E+09,9E+09,9E+09]];
    CONST robtarget Target_6550:=[[91.270074774,126.712231733,0],[0.882142515,0,0,-0.470982573],[0,0,0,0],[9E+09,9E+09,9E+09,9E+09,9E+09,9E+09]];
    CONST robtarget Target_6560:=[[84.332416711,119.042831364,0],[0.882142515,0,0,-0.470982573],[0,0,0,0],[9E+09,9E+09,9E+09,9E+09,9E+09,9E+09]];
    CONST robtarget Target_6570:=[[84.332416711,117.523771388,0],[0.882142515,0,0,-0.470982573],[0,0,0,0],[9E+09,9E+09,9E+09,9E+09,9E+09,9E+09]];
    CONST robtarget Target_6580:=[[94.410082897,117.523771388,0],[0.882142515,0,0,-0.470982573],[0,0,0,0],[9E+09,9E+09,9E+09,9E+09,9E+09,9E+09]];
    CONST robtarget Target_6590:=[[94.410082897,112.42010037,0],[0.882142515,0,0,-0.470982573],[0,0,0,0],[9E+09,9E+09,9E+09,9E+09,9E+09,9E+09]];
    CONST robtarget Target_6600:=[[95.762416778,112.42010037,0],[0.882142515,0,0,-0.470982573],[0,0,0,0],[9E+09,9E+09,9E+09,9E+09,9E+09,9E+09]];
    CONST robtarget Target_6610:=[[95.762416778,119.042831364,0],[0.882142515,0,0,-0.470982573],[0,0,0,0],[9E+09,9E+09,9E+09,9E+09,9E+09,9E+09]];
    CONST robtarget Target_6620:=[[84.332416711,119.042831364,0],[0.882142515,0,0,-0.470982573],[0,0,0,0],[9E+09,9E+09,9E+09,9E+09,9E+09,9E+09]];
    CONST robtarget Target_6630:=[[95.762416778,111.225230022,0],[0.882142515,0,0,-0.470982573],[0,0,0,0],[9E+09,9E+09,9E+09,9E+09,9E+09,9E+09]];
    CONST robtarget Target_6640:=[[84.332416711,111.225230022,0],[0.882142515,0,0,-0.470982573],[0,0,0,0],[9E+09,9E+09,9E+09,9E+09,9E+09,9E+09]];
    CONST robtarget Target_6650:=[[84.332416711,104.07453306,0],[0.882142515,0,0,-0.470982573],[0,0,0,0],[9E+09,9E+09,9E+09,9E+09,9E+09,9E+09]];
    CONST robtarget Target_6660:=[[85.684750593,104.07453306,0],[0.882142515,0,0,-0.470982573],[0,0,0,0],[9E+09,9E+09,9E+09,9E+09,9E+09,9E+09]];
    CONST robtarget Target_6670:=[[85.684750593,109.706170046,0],[0.882142515,0,0,-0.470982573],[0,0,0,0],[9E+09,9E+09,9E+09,9E+09,9E+09,9E+09]];
    CONST robtarget Target_6680:=[[88.815496154,109.706170046,0],[0.882142515,0,0,-0.470982573],[0,0,0,0],[9E+09,9E+09,9E+09,9E+09,9E+09,9E+09]];
    CONST robtarget Target_6690:=[[88.815496154,104.454298054,0],[0.882142515,0,0,-0.470982573],[0,0,0,0],[9E+09,9E+09,9E+09,9E+09,9E+09,9E+09]];
    CONST robtarget Target_6700:=[[90.167830035,104.454298054,0],[0.882142515,0,0,-0.470982573],[0,0,0,0],[9E+09,9E+09,9E+09,9E+09,9E+09,9E+09]];
    CONST robtarget Target_6710:=[[90.167830035,109.706170046,0],[0.882142515,0,0,-0.470982573],[0,0,0,0],[9E+09,9E+09,9E+09,9E+09,9E+09,9E+09]];
